(* IEC 61131-3 sources: daoli-st-library/DL_Device (part 2) *)

(* ---- FB_DL_DeviceParamVerify.st ---- *)
(*==============================================================================
 * 组件名称 (Component)  : FB_DL_DeviceParamVerify
 * 所属子库 (Sublibrary) : DL_Device
 * 当前版本 (Version)    : 1.0.1
 * 兼容性   (Platform)   : CODESYS 3.5 / TwinCAT 3 / 汇川 InoProShop / Machine Expert
 *                         仅依赖 Standard.library（ABS / MAX / R_TRIG / TON）
 * 功能描述 (Function)   : 把「组态期望参数块」与「设备回读参数块」逐项按逐项容差比对，
 *                         给出差异项数、首个超差项下标、最大偏差与其下标，以及
 *                         「一致 / 不一致」结论。不一致结论锁存，须显式确认才清除。
 *                         现场用途：伺服与变频器换板、参数被误改后设备带着错参数运行，
 *                         人工翻参数页核几十项既慢又漏；上电自动核对能把「参数被改」
 *                         从一条偶发工艺异常变成一条明确报警。
 *                         回读未就绪约定：回读块全部为零视为「设备尚未回传」，
 *                         在回读超时窗内持续等待，超时即判故障；该约定写死在本件，
 *                         调用方若确有「全零合法」的参数块，须自行叠加就绪位后再调用。
 * 出口契约 (Exit)       : bVerified 为「本轮核对全部项在容差内」；bMismatch 为锁存结论，
 *                         由 bAcknowledge 上升沿清除；nDiffCount / fMaxDev 等明细在核对拍
 *                         刷新并在结论驻留相保持（HMI 可同时看到「锁存结论」与「最近明细」）；
 *                         bError 只由 030D / 030E / 030F 三码置位，bReset 上升沿统一清除。
 * 不内联姊妹件的理由    : 姊妹件 FC_DL_ArrayDiffSummary 是「统一容差」的通用双数组比对；
 *                         本件是「逐项容差 + 结论锁存 + 回读超时」的设备参数域件。若复用该函数，
 *                         逐项容差会被拆成最多 64 次函数调用，破坏「单拍内完成一次完整核对」
 *                         的一致性（每次调用之间的数组不可能被冻结），故本件自带单次遍历循环，
 *                         两次循环的职责并不重复：一个算差异摘要，一个判设备参数一致性并锁存。
 * 开源溯源 (Origin)     : 来源标签 codesys-forge-devicereader。许可证：该示例页面未显式声明
 *                         许可，按最严口径处置——零代码行复制、零注释引用、零结构体搬运。
 *                         借鉴点仅为「读出 → 比对 → 出报告」三段式流程骨架与函数域划分。
 *                         状态机、逐项容差回落规则、结论锁存、非有限值处置、码位全部自有，
 *                         clean-room 独立实现。
 * 码位说明 (Codes)      : 信息级 16#0003_014D（比对本数越界已钳位）/ 014E（核对一致）/
 *                         014F（负容差已取绝对值）；故障级 16#0003_030D（回读出现非有限值）/
 *                         030E（回读超时未就绪）/ 030F（非法相位兜底）。
 *                         共 6 码，全部落在 R12 计划第 1.2 节本件码段内。
 * 依赖     (Depends)    : 无 DL_ 内部依赖；Standard.library: ABS / MAX / R_TRIG / TON
 * 红线自检 (Redline)    : 1 ✓ 零全局变量表依赖、零外部变量声明、零物理地址
 *                         2 ✓ 纯 IEC 61131-3，无指针、无厂商库
 *                         3 ✓ 数组先判界（遍历上界取钳位后的项数）、容差先收敛到正数、
 *                             非有限值前置拦截、循环带守卫、超时仅在等待相计时
 *                         4 ✓ 全变量中英双语同行注释
 *                         5 ✓ 六态 ENUM + CASE 全覆盖 + ELSE 兜底（030F）
 *                         6 ✓ R_TRIG / TON 实例在 CASE 之外每拍无条件刷新
 *                         7 ✓ END_FUNCTION_BLOCK 位于文件最后有效行
 * 修订历史 (Revision)   :
 *   2026-11-15  v1.0.0  首版入库（R12 · Level 1 DL_Device 参数域校验）
 *   2026-11-15  v1.0.1  终审修复：事件码跨核对周期不清。原实现只在复位沿清 uErrorId，
 *                       一轮核对留下的 014E 会一直驻留：后续轮次的 014D / 014F 因「仅在
 *                       uErrorId 为零时置码」被永久压住，且不一致轮次里会出现「码说一致、
 *                       结论说不一致」。改为进入新一轮核对（空闲转等待）时清信息级码
 *============================================================================*)

(*-----------------------------------------------------------------------------
 * 枚举: E_DL_ParamVerifyPhase（归属 DL_Device，与本功能块同文件）
 * 含义: 参数核对流程的离散相位。步长留空位，便于后续插态。
 *----------------------------------------------------------------------------*)
TYPE E_DL_ParamVerifyPhase :
(
    eIdle      := 0,     // 空闲：等待使能 / Idle: waiting for enable
    eWaiting   := 10,    // 等待：等设备回读就绪，同时跑回读超时 / Waiting for the readback or the timeout
    eComparing := 20,    // 比对：单拍内完成全项遍历 / Comparing: one pass over every item in a single scan
    eMatch     := 30,    // 一致：结论驻留，等待复位 / Match: verdict held until reset
    eMismatch  := 40,    // 不一致：结论锁存，等待确认 / Mismatch: latched until acknowledged
    eFault     := 99     // 故障：回读非法或超时，等待复位 / Fault: bad readback or timeout
);
END_TYPE

(*-----------------------------------------------------------------------------
 * 结构体: ST_DL_ParamVerifyState（归属 DL_Device，与本功能块同文件）
 * 含义: 跨周期状态包，由调用方持有并在多台设备间独立维护。
 *----------------------------------------------------------------------------*)
TYPE ST_DL_ParamVerifyState :
STRUCT
    bLastVerdict  : BOOL;     // 上次核对结论，TRUE = 一致 / Last verdict, TRUE means consistent
    nLastDiffCount : INT;     // 上次超差项数 [项] / Last out of tolerance count
    nLastFirstIdx : INT;      // 上次首个超差项下标，0 = 无 [索引] / Last first offending index
    fLastMaxDev   : REAL;     // 上次最大绝对偏差 [工程单位] / Last maximum absolute deviation
    uVerifyCount  : UDINT;    // 累计核对次数 [次] / Accumulated verification count
END_STRUCT
END_TYPE

(*==============================================================================
 * 功能块: FB_DL_DeviceParamVerify
 * 调用约定: 每个扫描周期无条件调用一次；bEnable 为 FALSE 时相位与结论全部冻结。
 * 无状态泄漏: 除调用方持有的状态包外，全部状态驻留于实例私有 VAR，零全局引用。
 *============================================================================*)
FUNCTION_BLOCK FB_DL_DeviceParamVerify
VAR_INPUT
    bEnable       : BOOL;                        // 使能，FALSE 时结论与相位冻结 / Enable, freezes the verdict when FALSE
    bReset        : BOOL;                        // 上升沿复位故障与结论锁存 / Rising edge clears fault and verdict latch
    bAcknowledge  : BOOL;                        // 上升沿确认「不一致」结论 / Rising edge acknowledges a mismatch
    nItemCount    : INT := 1;                    // 比对本数 [项]，域 1~64 / Item count, 1..64
    afExpected    : ARRAY[1..64] OF REAL;        // 组态期望参数块 [工程单位] / Configured expectation block
    afActual      : ARRAY[1..64] OF REAL;        // 设备回读参数块 [工程单位] / Device readback block
    afTolerance   : ARRAY[1..64] OF REAL;        // 逐项容差 [工程单位]，0 或负值回落默认 / Per item tolerance
    fDefaultTol   : REAL := 0.01;                // 默认容差 [工程单位]，域不小于 1E-6 / Default tolerance
    tVerifyTimeout : TIME := T#5S;               // 回读超时 [毫秒]，零表示不监控 / Readback timeout, zero disables it
END_VAR
VAR_OUTPUT
    bVerified     : BOOL;                        // 全部项在容差内 TRUE / All items within tolerance
    bMismatch     : BOOL;                        // 不一致结论锁存，需确认 / Mismatch latched until acknowledged
    nDiffCount    : INT;                         // 超差项数 [项] / Out of tolerance item count
    nFirstDiffIdx : INT;                         // 首个超差项下标，0 = 无 [索引] / First offending index
    fMaxDev       : REAL;                        // 最大绝对偏差 [工程单位] / Maximum absolute deviation
    nMaxDevIdx    : INT;                         // 最大偏差下标，0 = 无 [索引] / Index of the maximum deviation
    bError        : BOOL;                        // 故障级锁存，仅 030D~030F 置位 / Latched fault
    uErrorId      : UDINT;                       // 事件码，0 = 无事件 / Event code, zero means none
    eState        : E_DL_ParamVerifyPhase;       // 主状态机当前相位 / Current phase
END_VAR
VAR_IN_OUT
    stVerify      : ST_DL_ParamVerifyState;      // 跨周期状态：上次结论与累计核对次数 / Persistent state bag
END_VAR
VAR
    fbTrigReset   : R_TRIG;                      // 复位沿，CASE 之外每拍刷新 / Reset edge, refreshed outside CASE
    fbTrigAck     : R_TRIG;                      // 确认沿，CASE 之外每拍刷新 / Acknowledge edge, refreshed outside CASE
    fbTimeout     : TON;                         // 回读超时，CASE 之外每拍刷新 / Readback timer, refreshed outside CASE
    ePhase        : E_DL_ParamVerifyPhase := E_DL_ParamVerifyPhase.eIdle;  // 内部相位 / Internal phase
    bInit         : BOOL := FALSE;               // 首扫标志，首扫不做任何比对 / First scan flag, no comparison on it
    nCountUse     : INT;                         // 生效比对本数 [项] / Effective item count
    fTolDef       : REAL;                        // 生效默认容差 [工程单位] / Effective default tolerance
    fTolUse       : REAL;                        // 单项生效容差 [工程单位] / Per item effective tolerance
    fDev          : REAL;                        // 单项绝对偏差 [工程单位] / Per item deviation
    fExp          : REAL;                        // 期望值快照 [工程单位] / Expected snapshot
    fAct          : REAL;                        // 回读值快照 [工程单位] / Actual snapshot
    bNonFinite    : BOOL;                        // 本轮出现非有限值 / Non finite value encountered
    bReadbackReady : BOOL;                       // 回读块已非全零 / Readback block is no longer all zero
    bAckUse       : BOOL;                        // 本轮确认沿快照 / Acknowledge edge snapshot
    nGuard        : DINT;                        // 循环守卫 / Loop guard
    i             : INT;                         // 遍历索引 [项] / Loop index
END_VAR
VAR CONSTANT
    DL_ITEM_MAX   : INT  := 64;                  // 项数上限，与数组维度一致 [项] / Item count ceiling
    DL_TOL_MIN    : REAL := 1.0E-6;              // 最小容差 [工程单位] / Minimum tolerance
    DL_ABS_MAX    : REAL := 1.0E30;              // 有限值判定上界 [工程单位] / Finite value bound
    DL_ZERO_EPS   : REAL := 1.0E-9;              // 回读就绪判零容差 [工程单位] / Readback zero tolerance
    DL_NO_TIMEOUT : TIME := T#0S;                // 超时关闭标记 [毫秒] / Timeout disabled marker
    DL_GUARD_MAX  : DINT := 128;                 // 循环守卫上限 [次] / Loop guard limit
END_VAR

(*------------------------------------------------------------------------------
 * 段 0｜边沿与定时器每拍无条件刷新（严禁放进 CASE 或 IF 内部）
 *      Edge instances and the timer refreshed unconditionally on every scan
 *-----------------------------------------------------------------------------*)
fbTrigReset(CLK := bReset);
fbTrigAck(CLK := bAcknowledge);
fbTimeout(IN := (ePhase = E_DL_ParamVerifyPhase.eWaiting) AND bEnable, PT := tVerifyTimeout);
bAckUse := fbTrigAck.Q;

(*------------------------------------------------------------------------------
 * 段 1｜首扫闸：未初始化的回读块全为零，直接比对会误判不一致，首扫只做初始化
 *      First scan gate: an uninitialised readback block would be misjudged
 *-----------------------------------------------------------------------------*)
IF NOT bInit THEN
    bInit  := TRUE;
    ePhase := E_DL_ParamVerifyPhase.eIdle;
    eState := ePhase;
    RETURN;
END_IF

(*------------------------------------------------------------------------------
 * 段 2｜复位沿：故障、结论锁存、事件码一次性清干净，相位回空闲
 *      Reset edge clears the fault, the latch and the event code in one go
 *-----------------------------------------------------------------------------*)
IF fbTrigReset.Q THEN
    bError    := FALSE;
    bMismatch := FALSE;
    bVerified := FALSE;
    uErrorId  := 16#0000_0000;
    ePhase    := E_DL_ParamVerifyPhase.eIdle;
END_IF

(*------------------------------------------------------------------------------
 * 段 3｜比对本数钳位：越界钳位后照常核对，只发信息码
 *      Item count clamp: clamp and keep verifying, informational only
 *-----------------------------------------------------------------------------*)
nCountUse := nItemCount;
IF nCountUse < 1 THEN
    nCountUse := 1;
    IF uErrorId = 16#0000_0000 THEN
        uErrorId := 16#0003_014D;
    END_IF
ELSIF nCountUse > DL_ITEM_MAX THEN
    nCountUse := DL_ITEM_MAX;
    IF uErrorId = 16#0000_0000 THEN
        uErrorId := 16#0003_014D;
    END_IF
END_IF

(*------------------------------------------------------------------------------
 * 段 4｜默认容差收敛：取绝对值后再抬到下限，非有限值一律落到下限
 *      Default tolerance: absolute value, floored to the minimum
 *-----------------------------------------------------------------------------*)
fTolDef := ABS(fDefaultTol);
IF NOT (fTolDef >= DL_TOL_MIN) THEN
    fTolDef := DL_TOL_MIN;
END_IF

(*------------------------------------------------------------------------------
 * 段 5｜主状态机：六态全覆盖 + ELSE 兜底
 *      Main state machine with every enum member and an ELSE fallback
 *-----------------------------------------------------------------------------*)
IF bEnable THEN

    CASE ePhase OF
        E_DL_ParamVerifyPhase.eIdle:
            (* 空闲转为等待：开新一轮核对，先清上一轮的信息级码，其余出口保持 *)
            (* Idle arms the wait phase and clears the previous cycle's info code *)
            uErrorId   := 16#0000_0000;     // 清陈旧信息级码（014E 若不清会压住本轮的 014D / 014F，并与本轮结论矛盾） / Clear the stale info code
            bNonFinite := FALSE;
            ePhase     := E_DL_ParamVerifyPhase.eWaiting;

        E_DL_ParamVerifyPhase.eWaiting:
            (* 就绪判据：回读块出现任何一个非零量即视为已回传 *)
            (* Readiness: any non zero value in the readback block counts as arrived *)
            bReadbackReady := FALSE;
            i              := 1;
            nGuard         := 0;
            WHILE (i <= nCountUse) AND (NOT bReadbackReady) AND (nGuard < DL_GUARD_MAX) DO
                nGuard := nGuard + 1;
                IF NOT (ABS(afActual[i]) <= DL_ZERO_EPS) THEN
                    bReadbackReady := TRUE;
                END_IF
                i := i + 1;
            END_WHILE;

            IF tVerifyTimeout = DL_NO_TIMEOUT THEN
                (* 调用方关闭超时监控：直接进入比对 *)
                (* Timeout monitoring disabled by the caller: go straight to comparing *)
                ePhase := E_DL_ParamVerifyPhase.eComparing;
            ELSIF fbTimeout.Q AND (NOT bReadbackReady) THEN
                bError    := TRUE;
                uErrorId  := 16#0003_030E;
                bVerified := FALSE;
                ePhase    := E_DL_ParamVerifyPhase.eFault;
            ELSIF bReadbackReady THEN
                ePhase := E_DL_ParamVerifyPhase.eComparing;
            END_IF

        E_DL_ParamVerifyPhase.eComparing:
            (* 单拍单次遍历：逐项容差、非有限值、首差、最大偏差一次算全 *)
            (* One pass computes tolerance fallback, non finite values, first and worst item *)
            nDiffCount    := 0;
            nFirstDiffIdx := 0;
            fMaxDev       := 0.0;
            nMaxDevIdx    := 0;
            bNonFinite    := FALSE;
            i             := 1;
            nGuard        := 0;

            WHILE (i <= nCountUse) AND (nGuard < DL_GUARD_MAX) DO
                nGuard := nGuard + 1;
                fExp   := afExpected[i];
                fAct   := afActual[i];

                (* 容差回落：负值取绝对值并留痕，零值回落默认，最后抬到下限 *)
                (* Tolerance fallback: absolute value, then default, then the floor *)
                fTolUse := afTolerance[i];
                IF fTolUse < 0.0 THEN
                    fTolUse := ABS(fTolUse);
                    IF uErrorId = 16#0000_0000 THEN
                        uErrorId := 16#0003_014F;
                    END_IF
                END_IF
                IF fTolUse <= 0.0 THEN
                    fTolUse := fTolDef;
                END_IF
                fTolUse := MAX(fTolUse, DL_TOL_MIN);

                IF NOT ((fExp >= -DL_ABS_MAX) AND (fExp <= DL_ABS_MAX))
                   OR NOT ((fAct >= -DL_ABS_MAX) AND (fAct <= DL_ABS_MAX)) THEN
                    (* 非有限值：该项计超差，且不参与最大偏差竞争（非数比较无意义）*)
                    (* Non finite: counted as a difference, excluded from the worst deviation *)
                    bNonFinite := TRUE;
                    nDiffCount := nDiffCount + 1;
                    IF nFirstDiffIdx = 0 THEN
                        nFirstDiffIdx := i;
                    END_IF
                ELSE
                    fDev := ABS(fExp - fAct);
                    IF fDev > fTolUse THEN
                        nDiffCount := nDiffCount + 1;
                        IF nFirstDiffIdx = 0 THEN
                            nFirstDiffIdx := i;
                        END_IF
                    END_IF
                    IF fDev > fMaxDev THEN
                        fMaxDev    := fDev;
                        nMaxDevIdx := i;
                    END_IF
                END_IF

                i := i + 1;
            END_WHILE;

            IF bNonFinite THEN
                (* 数据源已坏：锁故障，结论与明细同时落盘供取证 *)
                (* Broken data source: latch a fault and store the details for evidence *)
                bError    := TRUE;
                uErrorId  := 16#0003_030D;
                bVerified := FALSE;
                stVerify.bLastVerdict   := FALSE;
                stVerify.nLastDiffCount := nDiffCount;
                stVerify.nLastFirstIdx  := nFirstDiffIdx;
                stVerify.fLastMaxDev    := fMaxDev;
                ePhase := E_DL_ParamVerifyPhase.eFault;
            ELSIF nDiffCount = 0 THEN
                (* 一致：清锁存，累计次数只在进入一致相时加一 *)
                (* Match: clear the latch, the counter increments only on entry *)
                bVerified := TRUE;
                bMismatch := FALSE;
                IF uErrorId = 16#0000_0000 THEN
                    uErrorId := 16#0003_014E;
                END_IF
                stVerify.bLastVerdict   := TRUE;
                stVerify.nLastDiffCount := 0;
                stVerify.nLastFirstIdx  := 0;
                stVerify.fLastMaxDev    := 0.0;
                stVerify.uVerifyCount   := stVerify.uVerifyCount + 1;
                ePhase := E_DL_ParamVerifyPhase.eMatch;
            ELSE
                (* 不一致：结论锁存，明细随结论一同落盘 *)
                (* Mismatch: latch the verdict and store the details *)
                bVerified := FALSE;
                bMismatch := TRUE;
                stVerify.bLastVerdict   := FALSE;
                stVerify.nLastDiffCount := nDiffCount;
                stVerify.nLastFirstIdx  := nFirstDiffIdx;
                stVerify.fLastMaxDev    := fMaxDev;
                stVerify.uVerifyCount   := stVerify.uVerifyCount + 1;
                ePhase := E_DL_ParamVerifyPhase.eMismatch;
            END_IF

        E_DL_ParamVerifyPhase.eMatch:
            (* 一致相驻留：结论保持不变，只认复位沿（在段 2 统一处理）*)
            (* Match dwell: the verdict stays, only the reset edge leaves it *)
            bVerified := TRUE;
            bMismatch := FALSE;

        E_DL_ParamVerifyPhase.eMismatch:
            (* 不一致相驻留：锁存结论与明细，确认沿清除锁存并重新武装 *)
            (* Mismatch dwell: the latch is cleared by the acknowledge edge only *)
            bMismatch := TRUE;
            bVerified := FALSE;
            IF bAckUse THEN
                bMismatch := FALSE;
                ePhase    := E_DL_ParamVerifyPhase.eIdle;
            END_IF

        E_DL_ParamVerifyPhase.eFault:
            (* 故障相驻留：输出冻结，只认复位沿 *)
            (* Fault dwell: the outputs are frozen until the reset edge *)
            bError := TRUE;

        ELSE
            (* 兜底：枚举被在线改坏或跨版本不兼容，置终端安全态并锁存 *)
            (* Fallback: terminal safe state with the segment last code *)
            bError    := TRUE;
            uErrorId  := 16#0003_030F;
            bVerified := FALSE;
            ePhase    := E_DL_ParamVerifyPhase.eFault;
    END_CASE

END_IF

(*------------------------------------------------------------------------------
 * 段 6｜相位出口：内部相位镜像到出口引脚
 *      Phase mirror to the output pin
 *-----------------------------------------------------------------------------*)
eState := ePhase;
END_FUNCTION_BLOCK

(* ---- FB_DL_DualValveBlockSet.st ---- *)
(*
  ==================================================================
  组件名 Component  : FB_DL_DualValveBlockSet
  分类   Category   : DL_Device
  前缀   Naming     : FB_DL_ ｜ b/n/u/f/t/e/st 类型前缀制（R265）
  码位   Code ID    : 16#0003_072D（故障级：组态非法）｜ 16#0003_072E（故障级：
                      反馈不一致窗超时）
  版本   Version    : 1.0.1
  变更   CHANGELOG  : v1.0.1 tonMismatch 相位闸
  复杂度 Complexity  : 中
  功能   Purpose    : 双阀冗余块组控：双阀同令同闭（单指令源统一下发）+ 两路
                      位置反馈不一致窗判定（一阀卡滞 / 位置开关故障的启动期
                      与稳态期保护）；不一致持续超窗即锁存故障并切断指令出口。
  开源溯源 Origin    : 西门子 LBP（免费闭源）阀特性「命令-监视-判定」三段分层
                      组织方式借鉴（R26 沿用，只借骨不抄肉）；双阀不一致窗
                      判据与实现 clean-room，零代码复制。
  许可证 License    : MIT
  参考   Reference  : IEC 61131-3:2013 §6.6 状态机与 TON 语义；冗余阀组
                      「命令-监视-判定」公开工程组织口径
  平台   Platform   : 纯 IEC 61131-3（TON / R_TRIG / ENUM+CASE / 四则），三平台通用
  依赖   Depends    : 仅 Standard.library（TON / R_TRIG 属标准件）
  分工声明 Split     : FB_DL_SingleValveCtrl（单阀对象）/ FB_DL_ValvePairXor
                      （二取一表决）与本件互引；本件为「同令同闭 + 不一致窗」
                      冗余组控，表决逻辑归 ValvePairXor（R216）。
  归属 Ownership     : E_DL_DualValvePhase 属主为本文件（全库唯一定义，R264）；
                      引用件只引用不重声明。
  ------------------------------------------------------------------
  边界 Boundary     :
                      一 组态闸结构早退（族② 判据）：tMismatchWin ≤ 0 →
                         组态码 072D + 三件套 + RETURN（无浮点引脚，非有限
                         闸 N/A，本件域闸仅时限一项，逐项点名 R272）；
                      二 状态机 ENUM + CASE 必带 ELSE（非法态兜底落 eFault +
                         锁存 072D，禁静默）；本拍合法事件（指令沿 / 反馈
                         归队）优先于超时迁移（R275 同拍竞态）；
                      三 不一致窗口径：_bMismatch = (bFbValveA <> bFbValveB)
                         电平直比（BOOL 反馈无容差问题）；指令切换瞬态的不
                         一致由 tMismatchWin 吸收（窗时长须大于双阀响应差
                         上限，交付默认 T#10S，调用方改参须维持该配比）；
                         持续超窗 → 锁存 072E；
                      四 失败锁存 bMismatchFault + _bFaultLatch；锁存解除式
                         （可达自证，R152）：bResetCmd 上升沿清锁存回 eIdle
                         （输入引脚恒可达，无「置位即永久」路径）；
                      五 指令出口切断（安全语义）：bValveCmd = bOpenCmd AND
                         NOT _bFaultLatch AND bEnable——故障锁存 / 失能期间
                         指令出口强制 FALSE（双保险语义，切令不切监视）；
                      六 bEnable = FALSE 的语义写死（FB33-4 声明行）：强制
                         eIdle + 双出口复位（不 faults，使能断开 ≠ 阀组故障）；
                      七 TON / R_TRIG 段 0 无条件刷新（禁入分支，R7）；监视
                         TON IN 串故障锁存门控（FB50-1）；
                      八 首拍 _bInit 全量初始化；无全局、无外部变量、无物理
                         地址；无浮点量（全 BOOL / TIME / ENUM），无除法。
  错误码 Codes      :
    16#0003_072D【故障级】组态非法（tMismatchWin ≤ 0）或非法状态拦截（ELSE 兜底）
    16#0003_072E【故障级】两路位置反馈不一致持续超窗（tMismatchWin，疑似单阀
                         卡滞或位置开关故障）
  码位反证 Note     :
    072D 与 072E 不可合并：072D 与输入无关（组态即刻判，处置人 = 组态工程师），
    072E 需运行期反馈到达（处置人 = 现场阀检），可由场景还原（R90），分立。
  验收 Acceptance   :
    算法已证（脚本）：未跑 ｜ 编译器已证（三平台）：未跑
    V1 指令 ON + 双反馈同步 ON → bInSync、bValveCmd 跟随、无码
    V2 单反馈滞留超窗 → 锁存 072E、bValveCmd 切断、bMismatchFault
    V3 指令切换瞬态不一致 < 窗 → 不误报（窗吸收向量）
    V4 故障态 bResetCmd 上升沿 → 解锁回 eIdle（锁存解除可达向量）
    V5 tMismatchWin = T#0S → 组态早退 072D
    V6 失能 → eIdle + 双出口复位（不 faults）
    V7 非法枚举态（强改 eState）→ ELSE 兜底落 eFault + 072D
  修订记录 Revision  :
    2026-11-21  v1.0.0  R64 首版（批 3 · 序号 8，LBP 阀组组织方式 clean-room）
    2026-11-22  v1.0.1  R65 点修（tonMismatch 相位闸）：计时启动条件补 eRun
                        相位门控——仅运行监视相才累计不一致窗，非运行相强制
                        IN = FALSE（R300：计时启动与判定相不同源，修 v1.0.0
                        「eIdle 期反馈不一致已累计、迁入 eRun 即刻误触发
                        072E」的残留窗缺陷）；超时触发动作后窗残留由相位闸
                        + 锁存门控双路自清（本件无 _nStep 类步序量，窗残留
                        仅 tonMismatch 累计值），复位 / 重入不残留旧窗数据
  ==================================================================
*)
TYPE E_DL_DualValvePhase :
(
    eIdle  := 0,  // 待机：等指令 / idle, waiting for the command
    eRun   := 10, // 运行监视：指令生效，两路反馈一致窗监视 / the run phase with the mismatch window supervision
    eFault := 20  // 锁存故障：不一致超窗或非法态，复位沿解除 / a latched fault released by the reset edge
);
END_TYPE

FUNCTION_BLOCK FB_DL_DualValveBlockSet
VAR_INPUT
    bEnable     : BOOL := TRUE;   // 使能，FALSE 时强制 eIdle + 双出口复位（边界六）/ the enable, false forces the idle and resets both outlets
    bOpenCmd    : BOOL := FALSE;  // 开阀指令 [-]，双阀统一下发 / the open command issued to both valves
    bFbValveA   : BOOL := FALSE;  // 阀 A 位置反馈 [-] / the position feedback of the valve A
    bFbValveB   : BOOL := FALSE;  // 阀 B 位置反馈 [-] / the position feedback of the valve B
    bResetCmd   : BOOL := FALSE;  // 故障复位电平，上升沿清锁存回 eIdle（边界四解除式）/ the fault reset level, its rising edge releases the latch
    tMismatchWin: TIME := T#10S;  // 不一致监视窗 [毫秒]，须 > 0 且大于双阀响应差上限 / the mismatch window, positive and above the response spread
END_VAR
VAR_OUTPUT
    bValveCmd      : BOOL := FALSE;          // 阀组指令出口 [-]（故障 / 失能强制切断，边界五）/ the valve command outlet cut off on a fault or disable
    bInSync        : BOOL := FALSE;          // 双反馈同步 [-] / the two feedbacks in sync
    bMismatchFault : BOOL := FALSE;          // 不一致故障（锁存）[-] / the latched mismatch fault
    eState         : E_DL_DualValvePhase;    // 状态机出口 [状态] / the state machine outlet
    bValid         : BOOL := FALSE;          // 判据可用 [-] / the criteria are usable
    eErr           : UDINT := 16#0000_0000;  // 错误码，0 = 正常 / the error code, zero is ok
    bError         : BOOL := FALSE;          // 故障标志（故障级码同拍置位，R45 配对）/ the fault flag raised with a fault level code
END_VAR
VAR
    _bInit      : BOOL := FALSE;  // 首拍初始化标志（R310 / FB50-2）/ the first scan flag
    _eState     : E_DL_DualValvePhase := E_DL_DualValvePhase.eIdle; // 内部状态寄存器 / the internal state register
    _bFaultLatch: BOOL := FALSE;  // 故障锁存副本（仅复位沿清除）/ the fault latch copy
    _uLatch     : UDINT := 16#0000_0000; // 故障码锁存 [码]（复位沿清除，FB33-1）/ the latched fault code cleared by the reset edge
    _bMismatch  : BOOL := FALSE;  // 反馈不一致电平（逐拍重算）/ the mismatch level recomputed every scan
    _bCfgBad    : BOOL := FALSE;  // 组态非法标记（逐拍重算）/ the configuration fault flag
    rtReset     : R_TRIG;         // 复位沿实例，段 0 无条件刷新（R7）/ the reset edge instance refreshed unconditionally
    tonMismatch : TON;            // 不一致窗定时器，段 0 无条件刷新 / the mismatch window timer refreshed unconditionally
END_VAR  // R64 结构补齐：VAR 段缺失的 END_VAR（门禁机械修复）
VAR CONSTANT
    DL_DVP_TIME0 : TIME := T#0S;        // 时间零常量 [毫秒] / the time zero constant
    DL_DVP_ZEROU : UDINT := 16#0000_0000; // 码零常量 / the code zero constant
END_VAR

// 段 0｜定时器与沿检测无条件周期刷新（禁入分支，R7；监视 TON 串锁存门控，FB50-1）/ segment 0, the unconditional refresh
rtReset(CLK := bResetCmd); // 复位沿 / the reset edge
_bMismatch := (bFbValveA <> bFbValveB); // 不一致电平逐拍重算（BOOL 直比无容差问题）/ the mismatch level recomputed, a plain boolean compare
tonMismatch(IN := _bMismatch AND (NOT _bFaultLatch)
         AND (_eState = E_DL_DualValvePhase.eRun), PT := tMismatchWin); // 不一致窗计时（v1.0.1 相位闸：仅 eRun 运行监视相累计，非运行相强制 IN = FALSE；串锁存门控防复位同拍重锁；超时触发后相位 + 锁存双路使 IN 自清，窗累计零残留，复位 / 重入不残留旧窗）/ the mismatch window with the v1.0.1 phase gate, accumulated only in the run phase

// 段 1｜首拍初始化与复位沿作用域（R310 / R311）/ segment 1, the first scan init and the reset edge scope
IF NOT _bInit THEN // 首拍一拍 / the first scan
    _bInit := TRUE; // 置首拍标志 / raise the first scan flag
    _eState := E_DL_DualValvePhase.eIdle; // 状态显式落空闲 / place the state to idle
    _bFaultLatch := FALSE; // 故障锁存显式清零 / clear the fault latch explicitly
    _uLatch := DL_DVP_ZEROU; // 码锁存显式清零 / clear the latched code explicitly
END_IF
IF rtReset.Q THEN // 复位沿（作用域声明：清锁存 + 迁相位，R311）/ the reset edge with the declared scope
    _bFaultLatch := FALSE; // 清故障锁存（唯一解除路径，边界四自证可达）/ clear the fault latch, the only release path
    _uLatch := DL_DVP_ZEROU; // 清码锁存 / clear the latched code
    _eState := E_DL_DualValvePhase.eIdle; // 迁回空闲 / back to idle
END_IF

// 段 2｜组态域闸结构早退（边界一，族② 判据：tMismatchWin 逐项点名）/ segment 2, the structural early exit on an illegal configuration
_bCfgBad := (tMismatchWin <= DL_DVP_TIME0); // 组态非法（窗非正）/ an illegal configuration
IF _bCfgBad THEN // 组态非法：结构早退（出口三件套 + RETURN）/ an illegal configuration exits structurally
    eState := _eState; // 状态照实出口（冻结）/ export the state as is
    bValveCmd := FALSE; // 指令出口切断（组态非法期禁下发）/ cut the command outlet off
    bInSync := NOT _bMismatch; // 同步位照实 / the sync bit as is
    bMismatchFault := _bFaultLatch; // 故障锁存照实回放 / replay the latch
    bValid := FALSE; // 判据不可用 / the criteria are not usable
    eErr := 16#0003_072D; // 故障级：组态非法 / fault grade, an illegal configuration
    bError := TRUE; // 同拍置故障标志（R45 配对）/ raise the fault flag on the same scan
    RETURN; // 结构早退 / the structural early exit
END_IF

// 段 3｜失能分支：强制 eIdle + 双出口复位，不 faults（边界六声明行）/ segment 3, the disabled branch
IF NOT bEnable THEN // 失能 / disabled
    _eState := E_DL_DualValvePhase.eIdle; // 强制空闲 / force the idle
    _bFaultLatch := FALSE; // 锁存复位（使能断开 ≠ 阀组故障）/ clear the latch
    _uLatch := DL_DVP_ZEROU; // 码锁存复位 / clear the code
    eState := _eState; // 状态出口 / the state outlet
    bValveCmd := FALSE; // 指令出口复位 / the command outlet resets
    bInSync := FALSE; // 同步位复位（失能不声明同步）/ the sync bit resets
    bMismatchFault := FALSE; // 故障位复位 / the fault bit resets
    bValid := FALSE; // 失能即不可用 / the criteria are not usable while disabled
    bError := FALSE; // 失能不是故障 / a disabled device is not a fault
    eErr := DL_DVP_ZEROU; // 失能不发码 / no code is emitted while disabled
    RETURN; // 早退 / early return
END_IF

// 段 4｜主状态机（ENUM + CASE，ELSE 兜底；本拍事件优先于超时迁移，R275）/ segment 4, the main machine
CASE _eState OF
    E_DL_DualValvePhase.eIdle: // 空闲相 / the idle phase
        IF bOpenCmd AND (NOT _bFaultLatch) AND (NOT _bCfgBad) THEN // 指令电平 + 全量闸位复检（R274）/ the command with the full gate recheck
            _eState := E_DL_DualValvePhase.eRun; // 迁入运行监视相 / enter the run phase
        END_IF
    E_DL_DualValvePhase.eRun: // 运行监视相（本拍合法事件优先：反馈归队先消化，再消化超窗，R275）/ the run phase, the event before the timeout
        IF NOT bOpenCmd THEN // 事件优先：指令撤回 / the command withdrawn, the event goes first
            _eState := E_DL_DualValvePhase.eIdle; // 回空闲（监视件不锁运行态）/ back to idle
        ELSIF tonMismatch.Q THEN // 不一致持续超窗（卡滞 / 开关故障判据）/ the mismatch stayed through the window
            _bFaultLatch := TRUE; // 锁存故障 / latch the fault
            _uLatch := 16#0003_072E; // 故障级：不一致超窗 / fault grade, the mismatch through the window
            bError := TRUE; // 同拍置故障标志（R45 配对，段 6 故障分支沿用）/ raise the fault flag on the same scan
        END_IF
    E_DL_DualValvePhase.eFault: // 锁存故障相（驻留，解除由段 1 复位沿承担）/ the fault phase dwelling, the release belongs to the reset edge
        ; // 驻留语义由注释表达（禁自赋值死语句，R261）/ the dwell is expressed by this comment without a dead statement
    ELSE // 非法枚举值拦截（边界二：落故障相并锁存，禁静默）/ the illegal enumeration guard
        _bFaultLatch := TRUE; // 锁存故障 / latch the fault
        _uLatch := 16#0003_072D; // 故障级：非法状态拦截（归入组态族一码，出口同形，R90）/ fault grade, the illegal state in the configuration family
        bError := TRUE; // 同拍置故障标志（R45 配对）/ raise the fault flag on the same scan
        _eState := E_DL_DualValvePhase.eFault; // 落故障相 / force the fault phase
END_CASE

// 段 5｜故障锁存迁移闸（置于解除段之后防同拍抢迁，R258）/ segment 5, the latch to phase gate
IF _bFaultLatch AND (_eState <> E_DL_DualValvePhase.eFault) THEN // 已锁存但不在故障相 / latched outside the fault phase
    _eState := E_DL_DualValvePhase.eFault; // 迁入故障相 / enter the fault phase
END_IF

// 段 6｜统一出口（名实双出口同源，R191）/ segment 6, the unified outlet
eState := _eState; // 状态出口 / the state outlet
bValveCmd := bOpenCmd AND (NOT _bFaultLatch); // 指令出口与锁存同源切断（边界五安全语义）/ the command outlet cut off with the latch
bInSync := NOT _bMismatch; // 同步位与不一致电平同源取反 / the sync bit inverted from the mismatch level
bMismatchFault := _bFaultLatch; // 故障位与锁存同源 / the fault bit from the latch
bValid := NOT _bFaultLatch; // 判据可用（无锁存故障）/ usable without a latch
IF _bFaultLatch THEN // 故障锁存回放优先（不在故障相按当下输入重新推断，R152）/ the latched fault replays first
    bValid := FALSE; // 故障相不可用 / not usable in the fault phase
    bError := TRUE; // 故障位置位（R45 配对）/ raise the fault bit
    eErr := _uLatch; // 锁存码回放 / replay the latched code
ELSE // 无事件 / no event
    bError := FALSE; // 无故障 / no fault
    eErr := DL_DVP_ZEROU; // 正常 / ok
END_IF
END_FUNCTION_BLOCK

(* ---- FB_DL_EnergyMeterAccum.st ---- *)
(*==============================================================================
 * 组件名称 (Component)  : FB_DL_EnergyMeterAccum
 * 所属子库 (Sublibrary) : DL_Device
 * 当前版本 (Version)    : 1.0.1
 * 组件分类 (Category)   : 功能块（FUNCTION_BLOCK）· 能源计量 · 电表冻结值累计与需量
 * 兼容性   (Platform)   : CODESYS 3.5 / TwinCAT 3 / 汇川 InoProShop / Schneider
 *                         Machine Expert；纯 IEC 61131-3（第 3 版）语法，
 *                         仅依赖 Standard.library（R_TRIG / TON），无算术库依赖
 * 功能描述 (Function)   : 按电表冻结寄存器语义拼装 32 位电能累计值（正反向各一），
 *                         做单调性校验、换表与清零识别，并按窗口滑算平均需量与峰值
 *                         需量。输出正向、反向与净电能，以及换表次数、单拍换表脉冲。
 * 分层声明 (Layering)   : ① 本件只做「原始值拼装 + 累计 + 需量」，不做寄存器读取调度
 *                         （读取节拍归轮询主站件，本件由调用方按冻结值更新节拍调用）；
 *                         ② 不做分时电价、不做费率分段、不做报表归档；
 *                         ③ 字序入参复用 DL_MathData 既有枚举，不另立枚举、不重复声明。
 * 字序与字节序 (Order)  : 本件处理的是「字间序」——32 位电能由两个 16 位寄存器拼装，
 *                         厂家有的按高字在前、有的按低字在前；既有字节交换件处理的是
 *                         「字节内序」，两者层次不同、不可互相替代，参数切换时请勿混填。
 * 诊断分层 (Diagnosis)  : 遵循 NAMUR NE43「原始值域诊断与工程量分离」的原则：先判原始
 *                         32 位拼装值的单调性，再做工程量换算，诊断结论不依赖标定系数
 *                         ——标定系数填错只会让数值错，不会让「换表」判定失效。
 * 职责边界 (Scope)      : 不做 32 位回绕的无损续接（回绕按换表处理，属有意保守策略：
 *                         0.1 kWh 每 LSB 时满量程约 4.29 亿 kWh，真实场景回绕前必换表）。
 * 开源溯源 (Origin)     : 来源标签 namur-ne43。原创实现（参考 NAMUR NE43 的「原始值域
 *                         诊断与工程量分离」契约形态，以及电表冻结寄存器的工程惯例）。
 *                         仅借诊断分层的组织方式，拼装算法、单调性策略、窗口需量口径、
 *                         枚举、状态机与全部码位 100% 本库独立设计，clean-room 实现，
 *                         零代码行复制。NE43 为公开推荐规范（非代码），无代码复制问题。
 * 依赖     (Depends)    : E_DL_ByteOrder（DL_MathData 既有类型，本件只引用不声明）；
 *                         Standard.library: R_TRIG / TON
 * 故障码表 (Error codes):
 *   16#0003_0150【信息级】冻结值刷新抖动，差值在回退阈值内，保持上次累计不累加
 *   16#0003_0151【信息级】需量窗口小于 1 秒已按 1 秒兜底
 *   16#0003_0152【信息级】换表回退比例越界已钳到 0 至 1
 *   16#0003_0310【故障级】每 LSB 电能非正，量纲错且含除零隐患（锁存）
 *   16#0003_0311【故障级】有功功率非有限值，本拍不积分（锁存）
 *   16#0003_0312【故障级】非法状态兜底（锁存，终端安全态）
 * 码位占用 (Slot)       : 信息级 0150 / 0151 / 0152；故障级 0310 / 0311 / 0312。
 *                         全部落在 R12 本件分配块内，无跨块借用、无段外哨兵值。
 * 拍序纪律 (Cycle order) :
 *   ① ePhase     ：段 6 状态机（唯一位移点），段 8 复位分支是唯一回退点
 *   ② fImportAcc ：首拍基准装载 → 每拍单调性判定后单点写回；抖动拍保持不写
 *   ③ 窗口累加器 ：段 6 的采样分支累加，段 6 的窗口结算分支清零，两处互斥
 *   ④ uErrorId   ：段 9 单一优先级链，全拍只写一次
 * 需量口径 (Demand)     : 平均需量按「窗口内电能除以窗口秒数再乘 3600」折算为千瓦；
 *                         窗口长度取需量窗口参数，暂停期间窗口冻结、恢复后按剩余时间
 *                         续计（不重头），故暂停不会把需量摊薄。
 * 验收向量 (Acceptance) :
 *   V1 高位与低位拼装：高字 1、低字 16#86A0、每 LSB 0.1 → 原始 100000 → 正向 10000.0 kW 时
 *   V2 增量：下拍低字加 1 → 正向 10000.1、增量 0.1
 *   V3 换表：随后低字回 5 → 检出换表，单拍脉冲、换表次数 1、正向重载为 0.5 且无负增量
 *   V4 需量：有功 100 kW、窗口 15 分钟、满窗 → 平均需量 100.0、峰值 100.0
 *   V5 量纲错：每 LSB 为 0 → 故障位置位、码 0310
 * 偏离留档 (Deviation)  :
 *   ① 规格第 3.14 节的回退判据写成「低于累计值减去回退比例乘 32 位满量程乘标定系数」，
 *      该式与验收向量 V3 矛盾（满量程 4.29 亿 kWh 的 1% 远大于 10000.1，换表永远判不出）。
 *      本件改为「低于累计值乘（1 减回退比例）」，即按累计值的比例判定，与 V3 一致，
 *      也是现场对「回退比例」一词的通行理解。
 *   ② 规格要求「周期取窗口秒数除以拍数」，但首窗拍数未知。本件以常量化标称周期开窗，
 *      窗口结算时用实测拍数刷新估计值，并在头注释声明「必须放在固定周期任务中调用」。
 *   ③ 反向电能的换表不累加换表次数（次数只记正向表，避免一表两计）。
 *   ④ 规格 VAR 清单列有冻结沿实例，但本件没有与之配套的显示位输出，实例化后其输出
 *      无处消费即成为只置不用的死代码；故不实例化，bFreezePulse 引脚保留，累计逻辑
 *      每拍按原始值递推、与冻结脉冲无关（防止误把冻结沿当累加触发）。
 * 修订历史 (Revision)   :
 *   2026-11-15  v1.0.0  首版落盘（R12 · 泳道 C · 电能累计与需量件）
 *   2026-11-15  v1.0.1  终审修复：二次及以后的暂停会拉长需量窗口。原实现用「整窗减已用
 *                       时间」保存剩余时间，但恢复后定时器的预置值已是剩余窗，ET 属于该
 *                       剩余窗，两者相减把剩余时间算大（窗口 900 s、半程暂停两次会拉长到
 *                       约 1300 s），平均需量被摊薄。改为按本拍实际预置值（tPtUse）求差
 *============================================================================*)

(*------------------------------------------------------------------------------
 * 枚举: E_DL_MeterPhase（本块相位，归属本功能块并同文件发布）
 *       Phase enumeration owned by this block and published in the same file
 *-----------------------------------------------------------------------------*)
TYPE E_DL_MeterPhase :
(
    eIdle     := 0,   // 待机：参数闸门未过或未使能，输出保持 / Idle, parameters not yet accepted or disabled
    eSampling := 10,  // 采样：拼装、换算、单调性判定、窗口积分与需量结算 / Sampling, the whole accumulation path
    eHeld     := 20,  // 冻结：掉使能，窗口停在剩余时间处，输出保持 / Held, the window is parked at its remaining time
    eFault    := 99   // 故障：量纲错、功率非有限或非法状态，需复位退出 / Fault, needs a reset to leave
);
END_TYPE

(*------------------------------------------------------------------------------
 * 结构体: ST_DL_MeterState（跨周期状态，由调用方持有）
 *         Persistent state structure, owned by the caller
 *         说明：累计值、窗口累加器与换表计数必须跨周期保持，建议声明为保持型变量，
 *               否则重新上电会把窗口与峰值清空、并可能把首拍误判为换表
 *-----------------------------------------------------------------------------*)
TYPE ST_DL_MeterState :
STRUCT
    uImportPrev   : UDINT;      // 上次正向原始拼装值 [LSB] / Previous stitched import raw value
    uExportPrev   : UDINT;      // 上次反向原始拼装值 [LSB] / Previous stitched export raw value
    fImportAcc    : REAL;       // 正向累计电能 [kWh] / Accumulated import energy
    fExportAcc    : REAL;       // 反向累计电能 [kWh] / Accumulated export energy
    fWindowEnergy : REAL;       // 本窗口已积电能 [kWh] / Energy accumulated in the current window
    tWindowElapsed: TIME;       // 本窗口已用时间 [毫秒] / Elapsed time of the current window
    fDemandPeak   : REAL;       // 历史峰值需量 [kW]，仅复位可清 / Peak demand, cleared by reset only
    uResetCount   : UDINT;      // 换表与清零累计次数 [次] / Meter swap and clear counter
END_STRUCT
END_TYPE

FUNCTION_BLOCK FB_DL_EnergyMeterAccum
VAR_INPUT
    bEnable        : BOOL;                         // 使能，FALSE 时冻结累计与窗口 [-] / Enable, freezing accumulation and the window
    bReset         : BOOL;                         // 复位需量窗口与统计，上升沿有效 [-] / Rising edge resets the window statistics
    uImportHi      : UINT;                         // 正向有功电能高字 [LSB] / Import energy high word
    uImportLo      : UINT;                         // 正向有功电能低字 [LSB] / Import energy low word
    uExportHi      : UINT;                         // 反向有功电能高字 [LSB] / Export energy high word
    uExportLo      : UINT;                         // 反向有功电能低字 [LSB] / Export energy low word
    fActivePower   : REAL;                         // 当前有功功率 [kW] / Active power in kilowatts
    eWordOrder     : E_DL_ByteOrder := E_DL_ByteOrder.eAbcd; // 字序约定，复用既有枚举，默认大字序 [-] / Word order, defaults to the big word order
    fKwhPerLsb     : REAL := 0.1;                  // 每个 LSB 对应电能 [kWh/LSB]，域大于 0 / Kilowatt hours per LSB, must exceed zero
    tDemandWindow  : TIME := T#15M;                // 需量统计窗口 [毫秒]，域不小于 1 秒 / Demand window, at least one second
    fRegressRatio  : REAL := 0.01;                 // 判为换表的回退比例 [-]，域 0 到 1 / Regression ratio for a meter swap
    bFreezePulse   : BOOL;                         // 冻结寄存器刷新脉冲，仅用于显示锁存 [-] / Freeze register update pulse, display only
END_VAR
VAR_OUTPUT
    fImportTotal   : REAL;                         // 正向累计电能 [kWh] / Accumulated import energy
    fExportTotal   : REAL;                         // 反向累计电能 [kWh] / Accumulated export energy
    fNetTotal      : REAL;                         // 净电能，正向减反向 [kWh] / Net energy, import minus export
    fDemandAvg     : REAL;                         // 本窗口平均需量 [kW] / Average demand of the window
    fDemandPeak    : REAL;                         // 历史峰值需量 [kW]，由复位清零 / Peak demand, cleared by reset
    fWindowEnergy  : REAL;                         // 本窗口累计电能 [kWh] / Energy accumulated in the window
    bMeterReset    : BOOL;                         // 检到换表或清零，单拍脉冲 [-] / Meter swap detected, one-scan pulse
    uResetCount    : UDINT;                        // 换表与清零累计次数 [次] / Swap events counted
    bError         : BOOL;                         // 故障级锁存，仅 0310 0311 0312 置位 [-] / Latched fault, only fault level codes set it
    uErrorId       : UDINT;                        // 事件码，0 表示无事件 [代码] / Event code, zero means none
    eState         : E_DL_MeterPhase;              // 主状态机当前相位 [-] / Current phase of the main state machine
END_VAR
VAR_IN_OUT
    stMeter        : ST_DL_MeterState;             // 跨周期：上次原始值、累计基准、窗口累加器 [-] / Persistent raw values, accumulators and window state
END_VAR
VAR
    fbTrigReset    : R_TRIG;                       // 复位沿检测，主周期无条件刷新 [-] / Reset edge detector, refreshed unconditionally
    fbWindow       : TON;                          // 需量窗口计时，主周期无条件刷新 / Demand window timer, refreshed unconditionally
    ePhase         : E_DL_MeterPhase := E_DL_MeterPhase.eIdle; // 内部相位，对外经 eState 输出 [-] / Internal phase exported as eState
    bInit          : BOOL := FALSE;                // 首扫标志，初值 FALSE，判据取非 [-] / First-scan flag initialised FALSE
    bInitSync      : BOOL := FALSE;                // 累计基准已装载（首拍不产生增量）[-] / Accumulation baseline loaded flag
    bFaultLatch    : BOOL;                         // 故障锁存，仅复位分支清除 [-] / Fault latch, cleared by the reset path only
    uErrInt        : UDINT;                        // 故障级码寄存，锁存型 [代码] / Latched fault level code register
    uInfoCode      : UDINT;                        // 本拍信息级码，每拍重算 [代码] / Info level code recomputed every scan
    fLsbUse        : REAL := 1.0;                  // 生效每 LSB 电能 [kWh/LSB]，钳位后 / Effective kilowatt hours per LSB after clamping
    fRatioUse      : REAL := 0.01;                 // 生效回退比例 [-]，钳位后 / Effective regression ratio after clamping
    tWinUse        : TIME := T#15M;                // 生效窗口长度 [毫秒]，钳位后 / Effective window length after clamping
    tPtUse         : TIME := T#15M;                // 本拍窗口定时器预置值 [毫秒]，恢复模式取剩余时间 / Timer preset of this scan
    tRemain        : TIME := T#15M;                // 暂停时保存的窗口剩余时间 [毫秒] / Remaining window time saved on hold
    fWinSec        : REAL := 900.0;                // 窗口长度换算成秒 [秒] / Window length in seconds
    bWinRun        : BOOL;                         // 窗口定时器输入电平 [-] / Window timer input level
    bWinBreak      : BOOL;                         // 窗口定时器断输入一拍 [-] / One-scan break of the window timer
    bWinEnd        : BOOL;                         // 窗口到点标志 [-] / Window boundary flag
    bRestoreMode   : BOOL;                         // 恢复模式，定时器预置值取剩余时间 [-] / Restore mode, the timer uses the remaining time
    uImportRaw     : UDINT;                        // 正向电能 32 位拼装值 [LSB] / Stitched import raw value
    uExportRaw     : UDINT;                        // 反向电能 32 位拼装值 [LSB] / Stitched export raw value
    fImportNow     : REAL;                         // 本次正向电能换算值 [kWh] / Converted import value of this scan
    fExportNow     : REAL;                         // 本次反向电能换算值 [kWh] / Converted export value of this scan
    fRegressThr    : REAL;                         // 本拍回退判定阈值 [kWh] / Regression threshold of this scan
    nCycleCount    : DINT;                         // 本窗口累计拍数 [拍] / Scan counter of the current window
    fCycleEst      : REAL := 0.01;                 // 标称周期估计值 [秒] / Estimated nominal cycle in seconds
    eOrderAbcd     : E_DL_ByteOrder := E_DL_ByteOrder.eAbcd; // 字序比较基准：大字序口径（声明区取值，便于统一审查）[-] / Word order comparison baseline
    bSwap          : BOOL;                         // 本次判为换表或清零 [-] / Swap detected this scan
    bRegress       : BOOL;                         // 本次判为刷新抖动 [-] / Jitter detected this scan
    bPowerFinite   : BOOL;                         // 有功功率有限标志 [-] / Finite active power flag
END_VAR
VAR CONSTANT
    DL_MS_PER_SEC   : REAL := 1000.0;              // 每秒毫秒数 [毫秒] / Milliseconds per second
    DL_SEC_PER_HOUR : REAL := 3600.0;              // 每小时秒数 [秒] / Seconds per hour
    DL_EPS          : REAL := 1.0E-6;              // 浮点比较容差 [kWh] / Float comparison tolerance
    DL_LSB_FALLBACK : REAL := 1.0;                 // 每 LSB 电能非法时的兜底值 [kWh/LSB] / Fallback gain
    DL_PWR_MAX      : REAL := 1.0E9;               // 功率合理上限，超出视为非有限 [kW] / Power sanity limit
    DL_CYCLE_MIN    : REAL := 1.0E-3;              // 周期估计下限 [秒] / Lower cycle bound
    DL_CYCLE_MAX    : REAL := 1.0;                 // 周期估计上限 [秒] / Upper cycle bound
    DL_CYCLE_NOM    : REAL := 0.01;                // 首窗标称周期 [秒]，10 毫秒任务 / Nominal cycle for the first window
    DL_WIN_MIN      : TIME := T#1S;                // 窗口长度下限 [毫秒] / Minimum window length
    DL_TIME_ZERO    : TIME := T#0S;                // 时间零值基准 [毫秒] / Time zero reference
END_VAR

(*------------------------------------------------------------------------------
 * 段 1｜输出确定性默认值（单拍标志每拍预清零，R25 第一律）
 *      Deterministic defaults first, one-scan flags pre-cleared every scan
 *-----------------------------------------------------------------------------*)
bMeterReset  := FALSE;                          // 换表脉冲预清零（Swap pulse pre-cleared）
uInfoCode    := 16#0000_0000;                   // 信息级码每拍重算（Info code recomputed every scan）
bSwap        := FALSE;                          // 换表判定预清零（Swap verdict pre-cleared）
bRegress     := FALSE;                          // 抖动判定预清零（Jitter verdict pre-cleared）
bPowerFinite := FALSE;                          // 功率有限标志预清零（Finite power flag pre-cleared）

(*------------------------------------------------------------------------------
 * 段 2｜沿检测无条件刷新（红线：实例在 CASE 之外每拍必刷）
 *      Edge detection refreshed unconditionally outside the CASE
 *-----------------------------------------------------------------------------*)
fbTrigReset(CLK := bReset);

(*------------------------------------------------------------------------------
 * 段 3｜首扫初始化（唯一合法范式：初值 FALSE，判据取非）
 *      First-scan initialisation following the single legal pattern
 *-----------------------------------------------------------------------------*)
IF NOT bInit THEN
    stMeter.uImportPrev    := 0;                // 上次正向原始值清零（Previous import raw cleared）
    stMeter.uExportPrev    := 0;                // 上次反向原始值清零（Previous export raw cleared）
    stMeter.fImportAcc     := 0.0;              // 正向累计清零（Import accumulation cleared）
    stMeter.fExportAcc     := 0.0;              // 反向累计清零（Export accumulation cleared）
    stMeter.fWindowEnergy  := 0.0;              // 窗口累加器清零（Window accumulator cleared）
    stMeter.tWindowElapsed := DL_TIME_ZERO;     // 窗口已用时间清零（Window elapsed cleared）
    stMeter.fDemandPeak    := 0.0;              // 峰值需量清零（Peak demand cleared）
    stMeter.uResetCount    := 0;                // 换表次数清零（Swap counter cleared）
    nCycleCount            := 0;                // 窗口拍计数清零（Window scan counter cleared）
    fCycleEst              := DL_CYCLE_NOM;     // 周期估计取标称值（Cycle estimate set to the nominal value）
    fDemandAvg             := 0.0;              // 平均需量清零（Average demand cleared）
    bWinRun                := FALSE;            // 窗口定时器停（Window timer stopped）
    bRestoreMode           := FALSE;            // 恢复模式关闭（Restore mode off）
    bInitSync              := FALSE;            // 累计基准待装载（Baseline to be loaded）
    fLsbUse                := DL_LSB_FALLBACK;  // 生效增益先给兜底值（Effective gain pre-set to the fallback）
    fRatioUse              := 0.0;              // 生效回退比例先给零（Effective ratio pre-set to zero）
    tWinUse                := DL_WIN_MIN;       // 生效窗口先给下限（Effective window pre-set to the lower bound）
    ePhase                 := E_DL_MeterPhase.eIdle; // 相位复位为待机（Phase reset to idle）
    bInit                  := TRUE;             // 首扫只做一次（First scan runs once）
END_IF

(*------------------------------------------------------------------------------
 * 段 4｜参数闸门（量纲错属故障级，窗口与比例越界属信息级，只钳位不停机）
 *      Parameter gate, dimensional errors latch a fault while clamps stay informational
 *-----------------------------------------------------------------------------*)
IF fKwhPerLsb <= DL_EPS THEN
    fLsbUse     := DL_LSB_FALLBACK;             // 量纲错：先给兜底增益避免本拍出现零乘（Fallback gain avoids a zero product）
    bFaultLatch := TRUE;                        // 锁故障（Latch the fault）
    uErrInt     := 16#0003_0310;                // 0310 每 LSB 电能非正（Non-positive energy per LSB）
ELSE
    fLsbUse := fKwhPerLsb;                      // 合法增益直通（Valid gain passed through）
END_IF

IF tDemandWindow < DL_WIN_MIN THEN
    tWinUse   := DL_WIN_MIN;                    // 小于 1 秒按 1 秒兜底，防需量除零（Clamped to one second to avoid a zero divisor）
    uInfoCode := 16#0003_0151;                  // 0151 窗口过短已兜底（Window too short, clamped）
ELSE
    tWinUse := tDemandWindow;                   // 合法窗口直通（Valid window passed through）
END_IF

IF fRegressRatio < 0.0 THEN
    fRatioUse := 0.0;                           // 负比例无意义：钳到 0（A negative ratio is clamped to zero）
    uInfoCode := 16#0003_0152;                  // 0152 比例越界已钳位（Ratio clamped）
ELSIF fRegressRatio > 1.0 THEN
    fRatioUse := 1.0;                           // 超 1 无意义：钳到 1（A ratio above one is clamped）
    uInfoCode := 16#0003_0152;                  // 0152 比例越界已钳位（Ratio clamped）
ELSE
    fRatioUse := fRegressRatio;                 // 合法比例直通（Valid ratio passed through）
END_IF

IF tWinUse > DL_TIME_ZERO THEN
    fWinSec := DINT_TO_REAL(TIME_TO_DINT(tWinUse)) / DL_MS_PER_SEC; // 窗口秒数，防除零由上限闸门保证（Seconds of the window）
ELSE
    fWinSec := 1.0;                             // 零窗口兜底为 1 秒（Zero window falls back to one second）
END_IF

(*------------------------------------------------------------------------------
 * 段 5｜32 位电能拼装（字间序，与字节内序件层次不同）
 *      Thirty-two bit energy stitching by word order
 *-----------------------------------------------------------------------------*)
IF eWordOrder = eOrderAbcd THEN
    uImportRaw := SHL(UINT_TO_UDINT(uImportHi), 16) OR UINT_TO_UDINT(uImportLo); // 高字在前（High word first）
    uExportRaw := SHL(UINT_TO_UDINT(uExportHi), 16) OR UINT_TO_UDINT(uExportLo); // 高字在前（High word first）
ELSE
    uImportRaw := SHL(UINT_TO_UDINT(uImportLo), 16) OR UINT_TO_UDINT(uImportHi); // 低字在前（Low word first）
    uExportRaw := SHL(UINT_TO_UDINT(uExportLo), 16) OR UINT_TO_UDINT(uExportHi); // 低字在前（Low word first）
END_IF
fImportNow := UDINT_TO_REAL(uImportRaw) * fLsbUse; // 正向工程量换算（Import engineering conversion）
fExportNow := UDINT_TO_REAL(uExportRaw) * fLsbUse; // 反向工程量换算（Export engineering conversion）

(*------------------------------------------------------------------------------
 * 段 6｜窗口计时（无条件刷新；入口电平取上一拍状态，断输入一拍重启）
 *      Window timer refreshed unconditionally, restarted by a one-scan break
 *-----------------------------------------------------------------------------*)
IF bRestoreMode THEN
    tPtUse := tRemain;                          // 恢复模式用剩余时间作预置值（Restore mode uses the remaining time）
ELSE
    tPtUse := tWinUse;                          // 正常模式用整窗作预置值（Normal mode uses the full window）
END_IF
fbWindow(IN := bWinRun AND (NOT bWinBreak), PT := tPtUse);
bWinBreak := FALSE;                             // 断输入脉冲在实例调用后自清（Break pulse self-cleared after the call）
bWinEnd   := fbWindow.Q;                        // 到点标志在实例调用后取用（Boundary flag read after the call）
stMeter.tWindowElapsed := fbWindow.ET;          // 窗口已用时间转出（Elapsed time exported）

(*------------------------------------------------------------------------------
 * 段 7｜主状态机（枚举每个成员均有标签，末尾 ELSE 兜底到终端安全态）
 *      Main state machine, one label per member plus a trailing ELSE fallback
 *-----------------------------------------------------------------------------*)
CASE ePhase OF

    E_DL_MeterPhase.eIdle: // 待机：参数可用且使能后进入采样
        IF bFaultLatch THEN
            ePhase := E_DL_MeterPhase.eFault;   // 参数已锁故障：直接进故障态（Gate failed, enter the fault state）
        ELSIF bEnable THEN
            bWinRun := TRUE;                    // 启动窗口（Start the window）
            ePhase  := E_DL_MeterPhase.eSampling; // 进采样态（Enter the sampling state）
        END_IF

    E_DL_MeterPhase.eSampling: // 采样：单调性判定、窗口积分、需量结算
        bWinRun := TRUE;                        // 窗口持续计时（Window keeps timing）
        IF NOT bInitSync THEN
            stMeter.fImportAcc  := fImportNow;  // 首拍只装载基准，不产生增量（First scan loads the baseline only）
            stMeter.fExportAcc  := fExportNow;  // 首拍只装载基准（First scan loads the baseline only）
            stMeter.uImportPrev := uImportRaw;  // 首拍记录原始值（Raw value recorded on the first scan）
            stMeter.uExportPrev := uExportRaw;  // 首拍记录原始值（Raw value recorded on the first scan）
            bInitSync           := TRUE;        // 基准装载完成（Baseline loaded）
        ELSE
            (* 正向单调性：低于累计值乘（1 减回退比例）判换表，低于容差内判抖动 *)
            fRegressThr := stMeter.fImportAcc * (1.0 - fRatioUse); // 回退阈值按累计值比例给出（Threshold from the accumulated value）
            IF fImportNow < fRegressThr THEN
                bSwap := TRUE;                  // 先判：大幅回退，疑似换表或清零（Decide first, a large regression looks like a swap）
            ELSIF fImportNow < (stMeter.fImportAcc - DL_EPS) THEN
                bRegress := TRUE;               // 先判：小幅回退，疑似刷新抖动（Decide first, a small regression looks like jitter）
            END_IF
            IF bSwap THEN
                bMeterReset         := TRUE;    // 单拍换表脉冲（One-scan swap pulse）
                stMeter.uResetCount := stMeter.uResetCount + 1; // 换表次数累加（Swap counter incremented）
                stMeter.fImportAcc  := fImportNow; // 基准重载，不回填负增量（Baseline reloaded, never a negative increment）
            ELSIF bRegress THEN
                uInfoCode := 16#0003_0150;      // 0150 冻结值刷新抖动（Freeze refresh jitter）
            ELSE
                stMeter.fImportAcc := fImportNow; // 正常递推（Normal accumulation）
            END_IF
            (* 反向单调性：只做基准重载，不重复计入换表次数 *)
            fRegressThr := stMeter.fExportAcc * (1.0 - fRatioUse); // 反向回退阈值（Export threshold）
            IF fExportNow < fRegressThr THEN
                stMeter.fExportAcc := fExportNow; // 反向换表：基准重载（Export baseline reloaded）
            ELSIF fExportNow >= stMeter.fExportAcc THEN
                stMeter.fExportAcc := fExportNow; // 正常递推（Normal accumulation）
            END_IF
            stMeter.uImportPrev := uImportRaw;  // 记录本拍原始值（Record the raw value of this scan）
            stMeter.uExportPrev := uExportRaw;  // 记录本拍原始值（Record the raw value of this scan）
        END_IF
        (* 有功功率有限性闸门：非有限值本拍不积分，并锁故障 *)
        IF (fActivePower <> fActivePower) OR (ABS(fActivePower) > DL_PWR_MAX) THEN
            bPowerFinite := FALSE;              // 判为非法功率（Marked as invalid power）
            IF NOT bFaultLatch THEN
                bFaultLatch := TRUE;            // 只在无更早故障时锁存，保留首出码 / Latch only when no earlier fault exists
                uErrInt     := 16#0003_0311;    // 0311 有功功率非有限（Non-finite active power）
            END_IF
        ELSE
            bPowerFinite := TRUE;               // 判为合法功率（Marked as valid power）
        END_IF
        (* 窗口积分：仅合法功率参与，故障拍不污染窗口 *)
        IF bPowerFinite THEN
            stMeter.fWindowEnergy := stMeter.fWindowEnergy + (fActivePower * fCycleEst); // 电能累加，千瓦乘小时（Energy in kilowatt hours）
            nCycleCount           := nCycleCount + 1; // 窗口拍数累加（Window scan counter incremented）
        END_IF
        (* 窗口结算：平均需量、峰值需量、周期估计刷新、累加器清零 *)
        IF bWinEnd THEN
            IF fWinSec > DL_EPS THEN
                fDemandAvg := stMeter.fWindowEnergy / fWinSec * DL_SEC_PER_HOUR; // 千瓦时转千瓦（Kilowatt hours to kilowatts）
            END_IF
            IF fDemandAvg > stMeter.fDemandPeak THEN
                stMeter.fDemandPeak := fDemandAvg; // 峰值取大（Peak takes the larger value）
            END_IF
            IF nCycleCount > 0 THEN
                fCycleEst := fWinSec / DINT_TO_REAL(nCycleCount); // 用实测拍数刷新周期估计（Cycle estimate refreshed from the measured count）
                fCycleEst := LIMIT(DL_CYCLE_MIN, fCycleEst, DL_CYCLE_MAX); // 周期估计钳位（Cycle estimate clamped）
            END_IF
            stMeter.fWindowEnergy := 0.0;       // 窗口累加器清零（Window accumulator cleared）
            nCycleCount           := 0;         // 窗口拍数清零（Window scan counter cleared）
            bRestoreMode          := FALSE;     // 退出恢复模式（Leave restore mode）
            bWinBreak             := TRUE;      // 定时器断输入一拍后重启（Restart the timer after a one-scan break）
        END_IF
        IF NOT bEnable THEN
            tRemain      := tPtUse - fbWindow.ET; // 保存剩余时间：按本拍实际预置值算，恢复态取剩余窗而非整窗（Remaining time from the preset in force）
            IF tRemain < DL_WIN_MIN THEN
                tRemain := DL_WIN_MIN;          // 剩余时间下限兜底（Remaining time lower bound）
            END_IF
            bWinRun     := FALSE;               // 窗口停止推进（Window stops advancing）
            ePhase      := E_DL_MeterPhase.eHeld; // 进冻结态（Enter the held state）
        ELSIF bFaultLatch THEN
            ePhase := E_DL_MeterPhase.eFault;   // 功率非法：进故障态（Invalid power, enter the fault state）
        END_IF

    E_DL_MeterPhase.eHeld: // 冻结：输出保持，恢复后按剩余时间续计，不重头
        bWinRun := FALSE;                       // 冻结期间窗口不推进（The window does not advance while held）
        IF bEnable THEN
            bRestoreMode := TRUE;               // 进入恢复模式（Enter restore mode）
            bWinBreak    := TRUE;               // 定时器断输入一拍后按剩余时间重启（Restart with the remaining time）
            bWinRun      := TRUE;               // 窗口重新推进（The window advances again）
            ePhase       := E_DL_MeterPhase.eSampling; // 回采样态（Back to sampling）
        END_IF

    E_DL_MeterPhase.eFault: // 故障：输出保持，等复位沿（Fault, outputs held until the reset edge）
        bWinRun := FALSE;                       // 故障期间窗口停止（The window stops during a fault）

    ELSE
        bFaultLatch := TRUE;                    // 非法状态兜底锁存（Illegal state latched）
        uErrInt     := 16#0003_0312;            // 0312 非法状态兜底（Illegal state fallback code）
        ePhase      := E_DL_MeterPhase.eFault;  // 进终端安全态（Enter the terminal safe state）
END_CASE

(*------------------------------------------------------------------------------
 * 段 8｜复位（清需量窗口与统计；累计值属电表自身读数，不清零）
 *      Reset clears the window statistics; the accumulated energy follows the meter
 *-----------------------------------------------------------------------------*)
IF fbTrigReset.Q THEN
    stMeter.fWindowEnergy := 0.0;               // 窗口累加器清零（Window accumulator cleared）
    stMeter.fDemandPeak   := 0.0;               // 峰值需量清零（Peak demand cleared）
    stMeter.uResetCount   := 0;                 // 换表次数清零（Swap counter cleared）
    fDemandAvg            := 0.0;               // 平均需量清零（Average demand cleared）
    nCycleCount           := 0;                 // 窗口拍数清零（Window scan counter cleared）
    bRestoreMode          := FALSE;             // 恢复模式关闭（Restore mode off）
    bWinBreak             := TRUE;              // 窗口定时器重启（Window timer restarted）
    bInitSync             := FALSE;             // 累计基准重装，复位后首拍不判换表（Baseline reloaded, no false swap after a reset）
    bFaultLatch           := FALSE;             // 清故障锁存（Clear the fault latch）
    uErrInt               := 16#0000_0000;      // 清故障码（Clear the fault code）
    IF ePhase = E_DL_MeterPhase.eFault THEN
        ePhase := E_DL_MeterPhase.eIdle;        // 故障态复位回待机（Fault returns to idle）
    END_IF
END_IF

(*------------------------------------------------------------------------------
 * 段 9｜码位定级与出口（单一优先级链，全拍只写一次 uErrorId）
 *      Single priority chain and outlet mapping
 *-----------------------------------------------------------------------------*)
eState        := ePhase;                        // 相位出口（Phase outlet）
fImportTotal  := stMeter.fImportAcc;            // 正向累计出口（Import total outlet）
fExportTotal  := stMeter.fExportAcc;            // 反向累计出口（Export total outlet）
fNetTotal     := fImportTotal - fExportTotal;   // 净电能出口（Net energy outlet）
fWindowEnergy := stMeter.fWindowEnergy;         // 窗口电能出口（Window energy outlet）
fDemandPeak   := stMeter.fDemandPeak;           // 峰值需量出口（Peak demand outlet）
uResetCount   := stMeter.uResetCount;           // 换表次数出口（Swap counter outlet）

bError := bFaultLatch;                          // 故障位只反映故障级锁存（Fault bit reflects the latch only）
IF bError THEN
    uErrorId := uErrInt;                        // 故障级码优先透出（Fault level code has priority）
ELSE
    uErrorId := uInfoCode;                      // 无故障透出本拍信息级码（Info code exposed otherwise）
END_IF
END_FUNCTION_BLOCK

(* ---- FB_DL_FlowMeterKFactorDrift.st ---- *)
(*==============================================================================
 * 组件名称 (Component)  : FB_DL_FlowMeterKFactorDrift
 * 所属子库 (Sublibrary) : DL_Device
 * 当前版本 (Version)    : 1.0.2
 * 兼容性   (Platform)   : CODESYS 3.5 / TwinCAT 3 / 汇川 InoProShop / Machine Expert
 *                         仅依赖 Standard.library + DL_ 库内既有件，零厂商方言
 * 来源标签 (Source)     : roadmap-industry-pool-19.6（§19.6 已勾未注册漂移件重建，
 *                         本件为漂移修复件，收口时须同步补 registry 注册行）
 * 功能描述 (Function)   : 流量计 K 系数漂移核对：批次结算沿采样——
 *                         ① K 系数回读比对（委托 FB_DL_DeviceParamVerify 读-比-判）；
 *                         ② 批次总量比对（委托 FB_DL_FlowTotalizer 累计，基线总量对拍）；
 *                         ③ 漂移折算（委托 FC_DL_LinearScale 做总量占基线百分比）。
 *                         合成漂移率取两判据绝对值最大者分级：
 *                         达 fDriftWarnPct -> eMaintenanceReq；达 fDriftLimitPct ->
 *                         eOutOfSpec；组态故障 -> eFailure；未采样 -> eUnknown。
 * 委托清单 (Delegation) : FB_DL_DeviceParamVerify（DL_Device，读-比-判内核）
 *                         FB_DL_FlowTotalizer（DL_Process，批次累计内核）
 *                         FC_DL_LinearScale（DL_MathData，百分比折算内核）
 * 归属声明 (Ownership)  : E_DL_Ne107Status 归属 DL_Device\I_DL_DeviceHealth.st，
 *                         本件只引用不重声明（六态仲裁口径与 I_DL_DeviceHealth 对齐）。
 * 边界与语义披露 (Boundary disclosure) :
 *   1) 采样时机：仅批次结算沿（bBatchSettle 上升沿）采样，批次窗口未关闭不采样；
 *      结算沿拍读入当批累计量，下一拍才发内部清零脉冲（延迟一拍，防同拍读零）。
 *   2) 除零双闸：fKFactorBaseline <= 0 或 fBatchBaseline <= 0 组态级故障，不采样
 *      不折算（安全侧），锁存至复位沿 + 组态恢复。
 *   3) 漂移率非有限拦截：合成漂移过自反 + 差自减双判，非有限拒绝发布（不置
 *      eHealth 降级，保持上一有效分级），故障级码 + bError 三件套。
 *   4) 采样周期 tSample 仅作为 FlowTotalizer 的钳位判据基准注入，本件自身
 *      不做时间换算（<= T#0S 仍为组态非法）。
 *   5) K 比对语义受 DeviceParamVerify 六态状态机约束：回读流持续非零即连续核对，
 *      结算沿消费其最新结论；回读全零（等待相）视为「未取得结论」不判漂移。
 * 故障码表 (Error codes) :
 *   16#0003_0500 [故障级] K 基线 <= 0 或基线总量 <= 0（除零双闸），不采样
 *                 反证：不采样时 eHealth 恒 eUnknown，与「从未使能」组合相同，
 *                 码位是组态错误的唯一出口。
 *   16#0003_0501 [故障级] 采样周期组态非法（<= T#0S），不采样
 *                 反证：周期非法与基线非法都表现为不采样不分级，输出组合不可区分。
 *   16#0003_0502 [故障级] 漂移阈值组态非法（负值或 warn >= limit），不分级
 *                 反证：不分级时保持上一有效分级，与「阈值恰好未触及」组合
 *                 输出相同，无码不可区分。
 *   16#0003_0503 [故障级] 合成漂移率非有限，拒绝发布（保持上一有效分级）
 *                 反证：拒绝发布与「本批漂移恰好等于上批」输出组合相同。
 *   16#0003_0400 [信息级] 漂移达维护级（eMaintenanceReq 分级确认）
 *                 反证：eHealth 已表达分级，码位承载「本批采样触发了该分级」
 *                 事件事实供流水归档（分级是状态，码位是事件，二者不互代）。
 *   16#0003_0401 [信息级] 漂移达超规格级（eOutOfSpec 分级确认）
 *                 反证：与 0400 同理，且两码互异满足归因唯一（R190）。
 * 码位总账 (Code ledger) : 16#0003_0500 / 0501 / 0502 / 0503 用 ｜ 16#0003_0400 / 0401 用
 * 依赖     (Depends)    : FB_DL_DeviceParamVerify / FB_DL_FlowTotalizer / FC_DL_LinearScale
 * 红线自检 (Redline)    : R1 ✓ 零全局变量与 VAR_EXTERNAL ｜ R2 ✓ 零 %I/%Q 物理地址
 *                         R3 ✓ 纯 IEC 61131-3 + 库内委托件
 *                         R4 ✓ 除零双闸 / 非有限双判 / 域闸全枚举 / 码位 R45 配对
 *                         R5 ✓ 全变量中英双语同行注释 ｜ R6 ✓ 四态 ENUM + CASE + ELSE 兜底
 *                         R7 ✓ 一沿实例无条件刷新；被委托件每拍无条件调用
 * 修订历史 (Revision)   :
 *   2026-11-22  v1.0.0  首版入库（R68 构建轮 · 批 2 · 目标 6，§19.6 漂移件重建）
 *   2026-11-22  v1.0.1  终审就地修①：组态锁存解除路径可达化（复位沿 + 三项组态改对即清锁存，原 eFault 相不可达）
 *   2026-11-22  v1.0.2  R69 点修③：组态故障相实现 eHealth := eFailure（原 eFailure 仅声明未实现，
 *                       头注释「组态故障 -> eFailure」与实现不符；实现取「补分级」而非「改注释」）
 *============================================================================*)

(*-----------------------------------------------------------------------------
 * 枚举: E_DL_KDriftPhase（归属 DL_Device，与 FB_DL_FlowMeterKFactorDrift 同文件）
 *----------------------------------------------------------------------------*)
TYPE E_DL_KDriftPhase :
(
    eIdle    := 0,    // 未使能：不采样不分级 / Disabled, no sampling or grading
    eArmed   := 10,   // 已使能待结算沿：累计器在跑 / Armed, waiting for the settle edge
    eSampled := 20,   // 本批已采样并分级 / Batch sampled and graded
    eFault   := 99    // 组态故障锁存：拒绝采样 / Config fault latched, sampling refused
);
END_TYPE

(*==============================================================================
 * 功能块: FB_DL_FlowMeterKFactorDrift
 * 调用约定: 每个扫描周期无条件调用一次；bBatchSettle 为单拍沿语义。
 *============================================================================*)
FUNCTION_BLOCK FB_DL_FlowMeterKFactorDrift
VAR_INPUT
    fFlow           : REAL;                  // 瞬时流量 [L/min]，委托 Totalizer 累计 / Instantaneous flow [L per min]
    bBatchSettle    : BOOL;                  // 批次结算沿（上升沿 = 批次窗口关闭）/ Batch settle edge
    fKFactorBaseline: REAL := 1000.0;        // K 系数基线 [脉冲/L]，<= 0 组态非法 / K factor baseline [pulses per L]
    fKFactorReadback: REAL;                  // K 系数设备回读 [脉冲/L] / K factor device readback
    fKTolerance     : REAL := 0.02;          // K 比对容差 [脉冲/L] / K comparison tolerance
    fBatchBaseline  : REAL := 100.0;         // 批次基线总量 [L]，<= 0 组态非法 / Batch baseline total [L]
    fDriftWarnPct   : REAL := 2.0;           // 漂移维护级阈值 [%] / Drift maintenance threshold [%]
    fDriftLimitPct  : REAL := 5.0;           // 漂移超规格级阈值 [%] / Drift out-of-spec threshold [%]
    tSample         : TIME := T#1S;          // 采样周期基准 [ms]，注入 Totalizer / Sample period basis for the totalizer
    bEnable         : BOOL := TRUE;          // 使能 / Enable
    bReset          : BOOL;                  // 上升沿：清除组态故障锁存 / Rising edge: clear config latches
END_VAR
VAR_OUTPUT
    eHealth        : E_DL_Ne107Status;       // NE107 健康出口（六态，属主 I_DL_DeviceHealth）/ NE107 health verdict
    fDriftKPct     : REAL;                   // K 系数漂移率 [%] / K factor drift rate [%]
    fDriftBatchPct : REAL;                   // 批次总量漂移率 [%] / Batch total drift rate [%]
    fDriftPctEff   : REAL;                   // 合成漂移率（两判据绝对值最大）[%] / Combined drift, max magnitude
    bKMismatch     : BOOL;                   // K 回读超容差（读-比-判结论）/ K readback out of tolerance
    bSampled       : BOOL;                   // 本批采样脉冲（单拍）/ Batch sampled pulse, single scan
    bError         : BOOL;                   // 故障标志（组态类锁存）/ Fault flag, configuration class
    uErrorId       : UDINT;                  // 故障码，0 = 无故障 / Error code, 0 = none
    eState         : E_DL_KDriftPhase;       // 当前相位（供 HMI 诊断）/ Current phase for HMI diagnosis
END_VAR
VAR
    fbTrigSettle   : R_TRIG;                 // 结算沿检测实例 / Settle edge detector
    fbTrigReset    : R_TRIG;                 // 复位沿检测实例 / Reset edge detector
    fbTotal        : FB_DL_FlowTotalizer;    // 批次累计委托实例 / Batch totalizer delegate
    fbVerify       : FB_DL_DeviceParamVerify; // K 读-比-判委托实例 / K verify delegate
    stKVerify      : ST_DL_ParamVerifyState; // 委托件跨周期状态袋（VAR_IN_OUT 注入）/ Delegate state bag
    afKExp         : ARRAY[1..64] OF REAL;   // 委托件期望参数块（仅第 1 项使用）/ Delegate expectation block, item 1 only
    afKAct         : ARRAY[1..64] OF REAL;   // 委托件回读参数块（仅第 1 项使用）/ Delegate readback block, item 1 only
    afKTol         : ARRAY[1..64] OF REAL;   // 委托件容差块（仅第 1 项使用）/ Delegate tolerance block, item 1 only
    ePhaseInt      : E_DL_KDriftPhase;       // 主状态机内部当前态 / Internal state machine state
    bRstPend       : BOOL;                   // 延迟一拍的批次清零待发标志 / Delayed batch reset pending flag
    fBatchMeas     : REAL;                   // 结算沿采得的批次总量 [L] / Batch total sampled at settle
    bScaleOk       : BOOL;                   // 折算有效标志（LinearScale 出口）/ Scaling valid flag from LinearScale
    uScaleErr      : UDINT;                  // 折算错误码透传 / Scaling error code pass-through
    fDriftK        : REAL;                   // K 漂移率中间量 [%] / K drift intermediate
    fDriftBatch    : REAL;                   // 总量漂移率中间量 [%] / Batch drift intermediate
    fDriftEff      : REAL;                   // 合成漂移率中间量 [%] / Combined drift intermediate
    bCfgKBad       : BOOL;                   // K / 基线总量组态非法 / K or baseline config illegal
    bCfgTBad       : BOOL;                   // 采样周期组态非法 / Sample period illegal
    bCfgPBad       : BOOL;                   // 漂移阈值组态非法 / Drift thresholds illegal
    bFaultLatch    : BOOL;                   // 组态故障锁存（复位沿清除）/ Config fault latch, cleared by reset edge
    bKReady        : BOOL;                   // 委托件已取得 K 比对结论 / Delegate verdict available
    bSampledT      : BOOL;                   // 本拍采样脉冲内部副本 / Internal sampled pulse copy
    bErrorInt      : BOOL;                   // 本拍故障置位累加（出口归并）/ Fault set accumulator of this scan
    bFirstScan     : BOOL := TRUE;           // 上电首扫标志 / First-scan flag
END_VAR
VAR CONSTANT
    DL_KD_FIN_LIM  : REAL := 1.0E30;   // REAL 有限幅值判界 / REAL finiteness magnitude bound
    DL_KD_ITEM     : INT  := 1;        // 委托件比对本数 [项]，K 单项 / Delegate item count, single K item
END_VAR

(*------------------------------------------------------------------------------
 * 段 1｜无条件刷新区（红线 R7）：二沿 + 三委托件全部每拍调用，禁入分支
 *      Unconditional refresh: two edges and three delegates called every scan
 *-----------------------------------------------------------------------------*)
fbTrigSettle(CLK := bBatchSettle);
fbTrigReset(CLK := bReset);

(* 委托件引脚装配（仅第 1 项）：期望 = K 基线，实际 = K 回读 *)
(* Delegate pin wiring, item 1 only: expectation vs readback *)
afKExp[1] := fKFactorBaseline;
afKAct[1] := fKFactorReadback;
afKTol[1] := fKTolerance;

fbVerify(bEnable := bEnable, bReset := bReset, nItemCount := DL_KD_ITEM,
         afExpected := afKExp, afActual := afKAct, afTolerance := afKTol,
         stVerify := stKVerify);

fbTotal(fFlow := fFlow, bRstBatch := bRstPend, bEn := bEnable, tSample := tSample);

(* 延迟清零脉冲消化：上一结算拍置位的待发标志已随上调用发出，此处撤销 *)
(* Delayed reset pulse consumed: the pending flag went out with the call above *)
IF bRstPend THEN
    bRstPend := FALSE;
END_IF

(*------------------------------------------------------------------------------
 * 段 2｜上电首扫：相位与分级落安全侧
 *      First-scan init: phase and health verdict to the safe side
 *-----------------------------------------------------------------------------*)
IF bFirstScan THEN
    ePhaseInt      := E_DL_KDriftPhase.eIdle;
    eHealth        := E_DL_Ne107Status.eUnknown;
    bRstPend       := FALSE;
    fBatchMeas     := 0.0;
    fDriftK        := 0.0;
    fDriftBatch    := 0.0;
    fDriftEff      := 0.0;
    bFirstScan     := FALSE;
END_IF

(*------------------------------------------------------------------------------
 * 段 3｜每拍预清（FB32-1）：单拍标志，禁入锁存 / 快照
 *      Per-scan preset: single-scan flags only
 *-----------------------------------------------------------------------------*)
bErrorInt := FALSE;
bSampledT := FALSE;

(*------------------------------------------------------------------------------
 * 段 4｜组态域闸（R151 全枚举：基线双量 / 周期 / 阈值对，含非有限双判）
 *      Config gates: baselines, period, threshold pair, with non-finite checks
 *      解除路径（R152 自证）：复位沿 AND 全部组态非法条件消失
 *-----------------------------------------------------------------------------*)
bCfgKBad := (fKFactorBaseline <= 0.0) OR (fKFactorBaseline <> fKFactorBaseline)
            OR (fBatchBaseline <= 0.0) OR (fBatchBaseline <> fBatchBaseline)
            OR (ABS(fKFactorBaseline) >= DL_KD_FIN_LIM) OR (ABS(fBatchBaseline) >= DL_KD_FIN_LIM);
bCfgTBad := (tSample <= T#0S);
bCfgPBad := (fDriftWarnPct < 0.0) OR (fDriftLimitPct < 0.0)
            OR (fDriftWarnPct <> fDriftWarnPct) OR (fDriftLimitPct <> fDriftLimitPct)
            OR (fDriftWarnPct >= fDriftLimitPct);

IF bCfgKBad OR bCfgTBad OR bCfgPBad THEN
    bFaultLatch := TRUE;
END_IF

(* 终审就地修 v1.0.1（R68）：解除路径（R152 自证可达）——复位沿 AND 组态非法条件
 * 全部消失即清锁存。原实现把锁存清零只写在 eFault 相分支，而组态闸置锁存后
 * 并不迁相至 eFault（只回 eIdle / 驻留），eFault 相不可达 -> 锁存永不可解，
 * 组件保护/监视功能一次性永久失效直至 PLC 重启（终审两式①）。
 * Clear path made provably reachable: reset edge with the illegal config gone. *)
IF fbTrigReset.Q AND (NOT bCfgKBad) AND (NOT bCfgTBad) AND (NOT bCfgPBad) THEN
    bFaultLatch := FALSE;         // 锁存解除 / Latch cleared
    uErrorId    := 16#0000_0000;  // 码位随解除归零 / Code cleared with the latch
END_IF

IF bCfgKBad THEN
    uErrorId  := 16#0003_0500;   // 故障级：K / 基线总量非法 / Fault: K or baseline illegal
    bErrorInt := TRUE;
    eHealth   := E_DL_Ne107Status.eFailure;   // R69 点修③：故障级分级出口（原仅声明未实现）/ Fault-level verdict implemented
ELSIF bCfgTBad THEN
    uErrorId  := 16#0003_0501;   // 故障级：采样周期非法 / Fault: sample period illegal
    bErrorInt := TRUE;
    eHealth   := E_DL_Ne107Status.eFailure;   // R69 点修③：故障级分级出口 / Fault-level verdict
ELSIF bCfgPBad THEN
    uErrorId  := 16#0003_0502;   // 故障级：漂移阈值非法 / Fault: drift thresholds illegal
    bErrorInt := TRUE;
    eHealth   := E_DL_Ne107Status.eFailure;   // R69 点修③：故障级分级出口 / Fault-level verdict
END_IF

(* 组态锁存期健康出口保持最严等级：锁存未解除前不得回落（锁存回放，禁按当下输入重推，
 * R152 故障码锁存口径）。解除沿（复位沿 + 组态改对）后由下一结算沿重新分级。 *)
(* While latched the verdict stays at eFailure; it is only re-graded after the latch is cleared *)
IF bFaultLatch THEN
    eHealth := E_DL_Ne107Status.eFailure;     // 锁存期分级锁死最严 / Verdict pinned to failure while latched
END_IF

(*------------------------------------------------------------------------------
 * 段 5｜主状态机（红线 R6）：ENUM + CASE + ELSE 兜底
 *      Main state machine with the mandatory ELSE fallback
 *-----------------------------------------------------------------------------*)
CASE ePhaseInt OF

    E_DL_KDriftPhase.eIdle:
        IF bEnable AND (NOT bFaultLatch) THEN
            ePhaseInt := E_DL_KDriftPhase.eArmed;
        END_IF

    E_DL_KDriftPhase.eArmed:
        IF bFaultLatch OR (NOT bEnable) THEN
            ePhaseInt := E_DL_KDriftPhase.eIdle;
        ELSIF fbTrigSettle.Q THEN
            (* 结算沿采样：先读当批累计量，清零脉冲延迟一拍发出（防同拍读零） *)
            (* Settle edge: read the batch total first, delayed reset next scan *)
            fBatchMeas := fbTotal.fTotalBatch;
            bRstPend   := TRUE;
            bSampledT  := TRUE;
            ePhaseInt  := E_DL_KDriftPhase.eSampled;
        END_IF

    E_DL_KDriftPhase.eSampled:
        IF bFaultLatch OR (NOT bEnable) THEN
            ePhaseInt := E_DL_KDriftPhase.eIdle;
        ELSIF fbTrigSettle.Q THEN
            (* 连续批次：结算沿再次采样（累计器已在上一采样后清零重建） *)
            (* Consecutive batches: settle edge samples the rebuilt batch *)
            fBatchMeas := fbTotal.fTotalBatch;
            bRstPend   := TRUE;
            bSampledT  := TRUE;
        END_IF

    E_DL_KDriftPhase.eFault:
        IF fbTrigReset.Q AND (NOT bCfgKBad) AND (NOT bCfgTBad) AND (NOT bCfgPBad) THEN
            bFaultLatch := FALSE;          // 解除路径自证可达（R152）/ Clear path reachable
            uErrorId    := 16#0000_0000;
            ePhaseInt   := E_DL_KDriftPhase.eIdle;
        END_IF

    ELSE
        ePhaseInt := E_DL_KDriftPhase.eFault;
        uErrorId  := 16#0003_0500;
        bErrorInt := TRUE;

END_CASE;

(*------------------------------------------------------------------------------
 * 段 6｜采样拍折算（仅采样拍执行）：K 结论 + 总量百分比 + 合成分级
 *      Sample-scan folding: K verdict plus percent plus combined grading
 *-----------------------------------------------------------------------------*)
IF bSampledT THEN
    (* ① K 结论：委托件已取得比对结论才判漂移（等待相 = 未取得结论） *)
    bKReady    := fbVerify.bVerified OR fbVerify.bMismatch;
    bKMismatch := FALSE;
    fDriftK    := 0.0;
    IF bKReady THEN
        bKMismatch := fbVerify.bMismatch;
        IF fKFactorBaseline <> 0.0 THEN
            fDriftK := fbVerify.fMaxDev / fKFactorBaseline * 100.0;  // 除子已闸（0300 组态闸）/ Guarded divisor
        END_IF
    END_IF

    (* ② 总量漂移：委托 LinearScale 折算占基线百分比，再减 100 得漂移率 *)
    (* FC 直接调用 + 命名出口（库内惯例，见 FB_DL_RoomCo2DemandVent 先例） *)
    fDriftBatch := FC_DL_LinearScale(fIn := fBatchMeas,
                                     fInMin := 0.0,
                                     fInMax := fBatchBaseline,
                                     fOutMin := 0.0,
                                     fOutMax := 100.0,
                                     bClamp := FALSE,
                                     bValid => bScaleOk,
                                     uErrorId => uScaleErr) - 100.0;
    IF (NOT bScaleOk) OR (uScaleErr <> 16#0000_0000) THEN
        fDriftBatch := 0.0;      // 折算无效（基线组态闸已拦，此处兜底）/ Fold invalid, defensive zero
        uErrorId    := 16#0003_0500;
        bErrorInt   := TRUE;
    END_IF

    (* ③ 合成与分级：绝对值最大者承载，非有限拒绝发布（三件套 R258） *)
    fDriftEff := MAX(ABS(fDriftK), ABS(fDriftBatch));
    IF (fDriftEff <> fDriftEff) OR ((fDriftEff - fDriftEff) <> (fDriftEff - fDriftEff))
       OR (ABS(fDriftEff) >= DL_KD_FIN_LIM) THEN
        uErrorId  := 16#0003_0503;   // 故障级：合成漂移非有限 / Fault: combined drift non-finite
        bErrorInt := TRUE;
        (* 非有限拒绝发布：fDriftPctEff / eHealth 保持上一有效值（不写即保持） *)
        (* Non-finite: publish withheld, outputs hold the last valid values *)
    ELSE
        fDriftPctEff := fDriftEff;
        fDriftKPct     := fDriftK;
        fDriftBatchPct := fDriftBatch;
        IF fDriftEff >= fDriftLimitPct THEN
            eHealth   := E_DL_Ne107Status.eOutOfSpec;      // 超规格级 / Out of spec
            uErrorId  := 16#0003_0401;
        ELSIF fDriftEff >= fDriftWarnPct THEN
            eHealth   := E_DL_Ne107Status.eMaintenanceReq; // 维护级 / Maintenance required
            uErrorId  := 16#0003_0400;
        ELSE
            eHealth   := E_DL_Ne107Status.eOk;             // 在容差内 / Within tolerance
        END_IF
    END_IF
END_IF

(*------------------------------------------------------------------------------
 * 段 7｜输出单一出口（范式 P-05）
 *      Single output exit
 *-----------------------------------------------------------------------------*)
bSampled := bSampledT;   // 单拍脉冲统一出口（预清 + CASE 置位两段式）/ Unified single-scan exit
bError   := bErrorInt OR (ePhaseInt = E_DL_KDriftPhase.eFault);
eState   := ePhaseInt;
END_FUNCTION_BLOCK

(* ---- FB_DL_GripperForceVerify.st ---- *)
(*==============================================================================
 * 组件名称 (Component)  : FB_DL_GripperForceVerify
 * 所属子库 (Sublibrary) : DL_Device
 * 当前版本 (Version)    : 1.0.0
 * 兼容性   (Platform)   : CODESYS 3.5+ / TwinCAT 3 / 汇川 InoProShop / 施耐德 Machine Expert
 *                         仅依赖 Standard.library（TON / R_TRIG / ABS），零厂商私有库
 * 功能描述 (Function)   : 夹爪力窗判定——空夹 / 滑脱 / 超力三类特征判定，结果分档输出。
 *                         判定在"夹紧指令上升沿 → 验证窗结束"这一段内完成，三类特征用不同的
 *                         物理证据区分（这是本件的核心：三者混判会导致维护方向完全错误）：
 *                           ① **空夹**：整个验证窗内峰值力都没到 fForceLow —— 根本没夹到件
 *                              （或件不在位），属上料/定位问题；
 *                           ② **滑脱**：峰值曾达 fForceLow 以上，但窗末力已掉到 fForceLow 以下，
 *                              或窗内出现力衰减速率超过 fSlipRate 的快速下跌 —— 夹到了但滑了，
 *                              属夹爪面磨损/气压不足/件表面油污问题；
 *                           ③ **超力**：窗内峰值超过 fForceHigh —— 夹爪力过大，有压伤件的风险。
 *                         判定优先级：超力 > 滑脱 > 空夹 > 合格（超力是安全侧优先报）。
 *                         验证窗结束即出结论（eResult 分档），结论锁存到下一次夹紧指令或复位，
 *                         故 bOk 不会在窗口中途闪变。
 * 接口     (Interface)  : 输入 bGripCmd 夹紧指令、fForce 夹持力实测、fForceLow / fForceHigh 力窗
 *                         上下限（N）、fSlipRate 滑脱判定速率（N/s）、tVerify 验证窗（TIME）、
 *                         fVerifySec 同一窗的秒数值（REAL，与 tVerify 成对）、fDtS 采样周期（秒）、
 *                         bReset 复位；输出 eResult 判定结果、bOk 合格、bNg 不合格、fPeak 窗内
 *                         峰值力、fFellRate 窗内最大衰减速率、bVerified 结论已出、eState / eCause /
 *                         bError。
 * 边界     (Boundary)   : ① **属主边界（写死）：本件只判"夹持结果"，不控制夹爪电磁阀/伺服，
 *                         不做夹紧动作本身**。夹紧动作与到位属 `I_DL_Cylinder` / 夹爪执行件；
 *                         本件吃夹紧指令与力反馈，出判定结论供剔除与报警。
 *                         ② **PT 语义成对声明**：tVerify（TIME）与 fVerifySec（REAL）必须由调用方
 *                         成对给同一窗长。本件用 tVerify 驱动 TON，用 fVerifySec 参与速率换算
 *                         （fSlipRate × fVerifySec 的位移阈值思路相同），**全程不做 TIME→数值转换**。
 *                         ③ 组态闸：fForceLow <= 0.0、fForceHigh <= fForceLow、fSlipRate <= 0.0、
 *                         tVerify <= T#0S、fVerifySec <= eps、fDtS <= eps、任一 NaN → 故障锁存，
 *                         eResult 置 eFault 档（不宣称任何结论）。
 *                         ④ 单枚 TON（tonVerify）+ 两枚 R_TRIG（bGripCmd / bReset）段 0 无条件刷新；
 *                         tonVerify 用 IN :=（夹紧中 ∧ ¬Q）自复位，不靠外部沿清零（R188）。
 *                         ⑤ 故障相迁出唯一路径 = bReset 上升沿（R228B）。
 *                         ⑥ 零全局耦合（无 GVL / 无 VAR_EXTERNAL / 无物理地址）。
 * 分工声明 (Scope)      : 与 `FB_DL_AxisTorqueLimitGuard`（旋转轴力矩限）分工——那件是轴侧连续
 *                         力矩保护，本件是夹爪气动/电动夹持的**结果验证**；量程、时间尺度、
 *                         判据形态都不同，不可互替。
 * 来源标签 (Source Tag) : T2-6 ◐（开源参考：夹持力窗与滑脱判定特征参数域，零代码行复制）
 * 解除式   (Release)    : bReset 上升沿 ∧ 组态合法 → 清故障与结论，回等待相。
 *                         另：新的 bGripCmd 上升沿也会重开一次判定（正常工艺路径，非解除式）。
 * 码表     (Codes)      : 本件不占用任何全局数字码位。出口为 ENUM 结论分档 + BOOL 组；
 *                         数字码位待主控收口阶段统一派号。
 * 红线自检 (Redline)    : R1 ✓ 零 GVL/VAR_EXTERNAL ｜ R2 ✓ 零 %I/%Q/%M ｜ R3 ✓ 纯 IEC 61131-3
 *                         R4 ✓ 除零闸（fDtS）+ 力窗几何闸 + 浮点容差 ｜ R5 ✓ 声明逐行同行双语注释
 *                         R6 ✓ ENUM+CASE 含 ELSE ｜ R7 ✓ TON/R_TRIG 段 0 无条件刷新
 * 修订历史 (Revision)   : 2026-11-19  v1.0.0  R46 首版（批次 4 · 序号 18）
 *==============================================================================*)

TYPE E_DL_GfvResult :
(
    ePending  := 0,    // 验证窗进行中，结论未出 / Verification window in progress
    eOk       := 10,   // 合格（力在窗内且未滑脱） / Passed, force inside the window with no slip
    eEmpty    := 20,   // 空夹（峰值力从未达到下限） / Empty grip, peak never reached the lower limit
    eSlip     := 30,   // 滑脱（曾建立夹持力但掉出下限） / Slipped, grip established then lost
    eOverforce:= 40,   // 超力（峰值力超上限） / Over-force, peak exceeded the upper limit
    eFault    := 90    // 组态故障，未判定 / Configuration fault, not judged
);
END_TYPE

TYPE E_DL_GfvState :
(
    eIdle  := 0,    // 等待夹紧指令 / Awaiting a grip command
    eVerify:= 10,   // 验证窗进行相 / Verification window active
    eDone  := 20,   // 结论已出相（锁存） / Conclusion latched
    eFault := 90    // 组态故障相 / Configuration fault phase
);
END_TYPE

TYPE E_DL_GfvCause :
(
    eNone       := 0,   // 无异常 / No anomaly
    eCfgIllegal := 1,   // 组态非法（力窗倒置/速率非正/窗长非正/非有限） / Illegal configuration
    eEmptyGrip  := 2,   // 空夹 / Empty grip
    eSlipped    := 3,   // 滑脱 / Slipped
    eOverForce  := 4,   // 超力 / Over-force
    ePhaseBad   := 5    // 非法相位兜底 / Illegal phase fallback
);
END_TYPE

FUNCTION_BLOCK FB_DL_GripperForceVerify
VAR_INPUT
    bGripCmd    : BOOL := FALSE;        // 夹紧指令，上升沿开启验证窗 [-] / Grip command, rising edge opens the window
    fForce      : REAL := 0.0;          // 夹持力实测 [N] / Measured grip force [N]
    fForceLow   : REAL := 10.0;         // 力窗下限，域 > 0.0 [N] / Force window lower limit, > 0.0 [N]
    fForceHigh  : REAL := 80.0;         // 力窗上限，域 > fForceLow [N] / Force window upper limit, > lower [N]
    fSlipRate   : REAL := 50.0;         // 滑脱判定衰减速率，域 > 0.0 [N/s] / Slip decay rate threshold, > 0.0 [N/s]
    tVerify     : TIME := T#300MS;      // 验证窗时长（TIME 侧），域 > T#0S [ms] / Verification window, TIME side [ms]
    fVerifySec  : REAL := 0.3;          // 同一窗的秒数值（REAL 侧），域 > eps [s] / Same window in seconds, REAL side [s]
    fDtS        : REAL := 0.001;        // 采样周期，域 > eps [s] / Sample period, > eps [s]
    bReset      : BOOL := FALSE;        // 复位，上升沿清结论与故障 [-] / Reset, rising edge clears result and fault
END_VAR
VAR_OUTPUT
    eResult   : E_DL_GfvResult;     // 判定结果分档 [-] / Verdict grade
    bOk       : BOOL;               // 合格 [-] / Passed
    bNg       : BOOL;               // 不合格（空夹/滑脱/超力任一） [-] / Failed, any of empty, slip or over-force
    fPeak     : REAL;               // 窗内峰值力 [N] / Peak force inside the window [N]
    fFellRate : REAL;               // 窗内最大衰减速率（正数表示下跌） [N/s] / Maximum decay rate in the window, positive means falling [N/s]
    bVerified : BOOL;               // 结论已出（本件已判定，非进行中） [-] / Verdict delivered
    eState    : E_DL_GfvState;      // 状态出口 [-] / State outlet
    eCause    : E_DL_GfvCause;      // 成因出口（R190 归因唯一） [-] / Cause outlet
    bError    : BOOL;               // 故障标志（组态非法或不合格） [-] / Error flag
END_VAR
VAR
    _eState  : E_DL_GfvState := E_DL_GfvState.eIdle;    // 内部相位（CASE 唯一写入目标） / Internal phase
    _eCause  : E_DL_GfvCause := E_DL_GfvCause.eNone;    // 成因锁存量 / Latched cause
    _eResult : E_DL_GfvResult := E_DL_GfvResult.ePending;    // 结论锁存量 / Latched verdict
    tonVerify: TON;                 // 验证窗计时（自复位），段 0 无条件调用 / Verification window, self-resetting
    rtGrip   : R_TRIG;              // 夹紧指令沿实例，段 0 无条件调用 / Grip edge instance
    rtReset  : R_TRIG;              // 复位沿实例，段 0 无条件调用 / Reset edge instance
    _fPeak   : REAL;                // 窗内峰值力（锁存量） [N] / Peak force in the window, latched [N]
    _fPrev   : REAL;                // 上拍力快照（锁存量） [N] / Previous force, latched [N]
    _fFell   : REAL;                // 窗内最大衰减速率（锁存量） [N/s] / Maximum decay rate, latched [N/s]
    _bSlipSeen : BOOL;              // 窗内已见滑脱特征（锁存量） / Slip feature seen in the window, latched
    _bFault  : BOOL;                // 组态故障锁存位（锁存量） / Latched configuration fault
    _bCfgBad : BOOL;                // 组态非法当拍量 [-] / Illegal configuration this scan
    _bNonFin : BOOL;                // 输入非有限当拍量 [-] / Non-finite input this scan
    _fRate   : REAL;                // 当拍力变化速率的负向幅值 [N/s] / Present decay rate magnitude [N/s]
END_VAR
VAR CONSTANT
    DL_GFV_EPS : REAL := 1.0E-9;    // 时间与速率判零容差 [无量纲] / Time and rate epsilon
END_VAR

(* —— 段 0：判据派生 + 三实例无条件周期刷新 —— *)
_bNonFin := (fForce <> fForce) OR (fForceLow <> fForceLow)                // NaN 自反判（判等禁令唯一例外） / NaN self-reflexive tests
         OR (fForceHigh <> fForceHigh) OR (fSlipRate <> fSlipRate)
         OR (fVerifySec <> fVerifySec) OR (fDtS <> fDtS);
_bCfgBad := (fForceLow <= 0.0) OR (fForceHigh <= fForceLow)               // 力窗几何闸 / Force-window geometry gate
         OR (fSlipRate <= 0.0) OR (tVerify <= T#0S)                       // 速率与窗长闸 / Rate and window gates
         OR (fVerifySec <= DL_GFV_EPS) OR (fDtS <= DL_GFV_EPS) OR _bNonFin;   // 成对秒值与非有限 / Paired seconds and non-finite
rtGrip(CLK := bGripCmd);                                                  // 夹紧沿，每拍必调（R228A） / Grip edge, every scan
rtReset(CLK := bReset);                                                   // 复位沿，每拍必调 / Reset edge, every scan
tonVerify(IN := (_eState = E_DL_GfvState.eVerify) AND (NOT tonVerify.Q), PT := tVerify);   // 验证窗，自复位（R188） / Verification window, self-resetting

(* —— 段 1：单拍量预清零（锁存量 _fPeak/_fFell/_bSlipSeen/_eResult/_bFault 不入清单） —— *)
bOk       := FALSE;     // 合格位预清 / Passed preset
bNg       := FALSE;     // 不合格位预清 / Failed preset
bVerified := FALSE;     // 结论已出位预清 / Verified preset
bError    := FALSE;     // 故障标志预清（R45 配对） / Error flag preset

(* —— 段 2：复位沿（清结论与故障，回等待相） —— *)
IF rtReset.Q THEN
    _bFault    := FALSE;                            // 清故障锁存 / Clear the fault latch
    _bSlipSeen := FALSE;                            // 清滑脱特征 / Clear the slip feature
    _fPeak     := 0.0;                              // 峰值清零 / Peak cleared
    _fFell     := 0.0;                              // 衰减速率清零 / Decay rate cleared
    _eCause    := E_DL_GfvCause.eNone;              // 清成因 / Clear cause
    _eResult   := E_DL_GfvResult.ePending;          // 结论回进行中位 / Verdict back to pending
    _eState    := E_DL_GfvState.eIdle;              // 回等待相（R228B 迁出路径） / Back to idle, the R228B exit
END_IF
IF _bCfgBad THEN
    _bFault  := TRUE;                               // 组态非法锁存 / Latch illegal configuration
    _eCause  := E_DL_GfvCause.eCfgIllegal;          // 归因：组态非法 / Cause: illegal configuration
    _eResult := E_DL_GfvResult.eFault;              // 结论置故障档（不宣称） / Verdict set to fault, nothing claimed
    _eState  := E_DL_GfvState.eFault;               // 入故障相 / Enter fault phase
END_IF

(* —— 段 3：夹紧沿开启新一次验证（工艺路径，不属解除式） —— *)
IF rtGrip.Q AND (NOT _bCfgBad) THEN
    _fPeak     := 0.0;                              // 峰值重置 / Peak reset
    _fFell     := 0.0;                              // 衰减速率重置 / Decay rate reset
    _bSlipSeen := FALSE;                            // 滑脱特征重置 / Slip feature reset
    _fPrev     := fForce;                           // 力快照对齐（防首拍伪速率） / Align the snapshot to avoid a spurious first-scan rate
    _eResult   := E_DL_GfvResult.ePending;          // 结论进行中 / Verdict pending
    _eState    := E_DL_GfvState.eVerify;            // 入验证相 / Enter the verification phase
END_IF

(* —— 段 4：验证窗内的峰值与衰减跟踪（单点写入锁存量，避免同拍抹除，R187） —— *)
IF (_eState = E_DL_GfvState.eVerify) AND (NOT _bCfgBad) THEN
    IF fForce > _fPeak THEN
        _fPeak := fForce;                                       // 峰值跟踪 / Track the peak
    END_IF
    _fRate := (_fPrev - fForce) / fDtS;                         // 衰减速率（正数=下跌），分母已闸 / Decay rate, denominator gated
    IF _fRate > _fFell THEN
        _fFell := _fRate;                                       // 记录窗内最大衰减速率 / Track the maximum decay rate
    END_IF
    IF (_fRate > fSlipRate) AND (_fPeak >= fForceLow) THEN
        _bSlipSeen := TRUE;                                     // 已达下限后快速下跌 = 滑脱特征 / Fast decay after reaching the limit means slip
    END_IF
    _fPrev := fForce;                                           // 力快照更新 / Update the snapshot
END_IF

(* —— 段 5：窗末判定（三类特征按 超力 > 滑脱 > 空夹 > 合格 的优先级） —— *)
IF (_eState = E_DL_GfvState.eVerify) AND tonVerify.Q AND (NOT _bCfgBad) THEN
    IF _fPeak > fForceHigh THEN
        _eResult := E_DL_GfvResult.eOverforce;                  // 超力（安全侧最高优先） / Over-force, highest priority
        _eCause  := E_DL_GfvCause.eOverForce;
    ELSIF _bSlipSeen OR ((_fPeak >= fForceLow) AND (fForce < fForceLow)) THEN
        _eResult := E_DL_GfvResult.eSlip;                       // 滑脱：曾达下限但已掉出 / Slipped: reached the limit then lost it
        _eCause  := E_DL_GfvCause.eSlipped;
    ELSIF _fPeak < fForceLow THEN
        _eResult := E_DL_GfvResult.eEmpty;                      // 空夹：峰值从未达下限 / Empty: peak never reached the limit
        _eCause  := E_DL_GfvCause.eEmptyGrip;
    ELSE
        _eResult := E_DL_GfvResult.eOk;                         // 合格 / Passed
        _eCause  := E_DL_GfvCause.eNone;
    END_IF
    _eState := E_DL_GfvState.eDone;                             // 结论相 / Verdict phase
END_IF

(* —— 段 6：锁存相位迁移闸 —— *)
IF _bFault AND (_eState <> E_DL_GfvState.eFault) THEN
    _eState := E_DL_GfvState.eFault;                            // 锁存即入故障相 / Latch enters fault phase
END_IF

(* —— 段 7：相位机（ENUM 全成员显式标签 + ELSE 兜底，R128） —— *)
CASE _eState OF

E_DL_GfvState.eIdle:
    IF _bCfgBad THEN                                            // 出口 1：组态非法 / Illegal configuration
        _eState := E_DL_GfvState.eFault;
    ELSIF rtGrip.Q THEN                                         // 出口 2：夹紧沿 / Grip edge
        _eState := E_DL_GfvState.eVerify;
    END_IF

E_DL_GfvState.eVerify:
    IF _bCfgBad THEN                                            // 出口 1：组态转非法 / Configuration went illegal
        _eState := E_DL_GfvState.eFault;
    ELSIF (_eResult <> E_DL_GfvResult.ePending) THEN            // 出口 2：结论已出 / Verdict delivered
        _eState := E_DL_GfvState.eDone;
    END_IF

E_DL_GfvState.eDone:
    IF _bCfgBad THEN                                            // 出口 1：组态转非法 / Configuration went illegal
        _eState := E_DL_GfvState.eFault;
    ELSIF rtGrip.Q THEN                                         // 出口 2：新一次夹紧 / A new grip
        _eState := E_DL_GfvState.eVerify;
    ELSIF rtReset.Q THEN                                        // 出口 3：复位回等待相 / Reset back to idle
        _eState := E_DL_GfvState.eIdle;
    END_IF

E_DL_GfvState.eFault:
    IF rtReset.Q AND (NOT _bCfgBad) THEN                        // 出口：复位且组态已合法才迁出（R228B） / Reset with legal config
        _eState := E_DL_GfvState.eIdle;
    END_IF

ELSE
    _eCause  := E_DL_GfvCause.ePhaseBad;                        // 归因：非法相位 / Cause: illegal phase
    _eState  := E_DL_GfvState.eFault;                           // 强拉故障相 / Force fault phase
    _eResult := E_DL_GfvResult.eFault;                          // 结论置故障档 / Verdict to fault
    bError   := TRUE;                                           // 故障标志 / Error flag

END_CASE

(* —— 段 8：出口单点映射（结论分档与 bOk/bNg 同源；名实双出口，R191） —— *)
eResult   := _eResult;                                          // 结论出口 / Verdict outlet
fPeak     := _fPeak;                                            // 峰值出口 / Peak outlet
fFellRate := _fFell;                                            // 衰减速率出口 / Decay rate outlet
bVerified := (_eResult <> E_DL_GfvResult.ePending) AND (_eResult <> E_DL_GfvResult.eFault);   // 已判定且非故障档 / Judged and not in the fault grade
bOk       := (_eResult = E_DL_GfvResult.eOk);                    // 合格 / Passed
bNg       := (_eResult = E_DL_GfvResult.eEmpty) OR (_eResult = E_DL_GfvResult.eSlip)
          OR (_eResult = E_DL_GfvResult.eOverforce);             // 三类不合格 / Any of the three failure types
bError    := _bFault OR bNg;                                     // 故障标志 = 组态故障或不合格 / Error = config fault or failed verdict
eState    := _eState;                                            // 状态出口 / State outlet
eCause    := _eCause;                                            // 成因出口 / Cause outlet

END_FUNCTION_BLOCK
